(* IEC 61131-3 sources: daoli-st-library/DL_MathData (part 5) *)

(* ---- FC_DL_SaturateIncr.st ---- *)
(*==============================================================================
 * 组件名称 (Component)  : FC_DL_SaturateIncr
 * 所属子库 (Sublibrary) : DL_MathData ｜ 版本 (Version) : 1.0.0 ｜ 2026-11-23
 * 兼容性   (Platform)   : CODESYS 3.5+ / TwinCAT 3 / 汇川 InoProShop / 施耐德 Machine Expert
 *                         仅依赖 IEC 61131-3 算术运算符与 ABS，零厂商私有库
 * 功能描述 (Function)   : 带上下限的原地递增饱和（FC 形态）：把 VAR_IN_OUT 引脚 fX 原地
 *                         +1.0（步进常量 DL_SINC_STEP），结果超上限 fMax 则饱和到 fMax，
 *                         低于下限 fMin 则抬升到 fMin。用于配方号 / 档位 / 索引游标类
 *                         计数递增，替代任何不经限位的裸 `x := x + 1`。
 *                         **原地语义**：写回点唯一（段 5），返回 FALSE 的所有出口均不写 fX，
 *                         保证「失败不推进」。
 * 接口     (Interface)  : VAR_IN_OUT fX 被递增的量（本件原地更新）[工程单位]；
 *                         输入 fMin 下限、fMax 上限（有效域 fMin ≤ fMax）[工程单位]；
 *                         输出 fY 递增后值（镜像 fX）[工程单位]、bSaturated 本拍是否饱和、
 *                         eErrCode（E_DL_SaturateErr）；返回值 = 递增已生效标志。
 * 边界     (Boundary)   : ① fMin > fMax → 故障级 eBadLimit，fX 不写回（保持原值）。
 *                         ② 任一入参非有限 → 故障级 eNonFinite，fX 不写回。
 *                         ③ fX + 1 溢出为非有限 → 故障级 eNonFinite，fX 不写回（不饱和猜测）。
 *                         ④ 上限饱和与下限抬升为两个独立分支、两个独立码值（R190 归因唯一）。
 *                         ⑤ 容差 DL_SINC_EPS（1E-6）用于「恰好等于限值」的判定，禁浮点判等。
 *                         ⑥ 零全局耦合（无 GVL / VAR_EXTERNAL / 物理地址）。
 * 码表     (Codes)      : 本件不占用全局数字码位（R297 零码位范式）；出口为 BOOL + LREAL +
 *                         本文件内 enum E_DL_SaturateErr（全库唯一属主，与递减件共用同族枚举）。
 * 分工声明 (Scope)      : 递减同族件为 FC_DL_SaturateDecr（共用 E_DL_SaturateErr）；
 *                         整数类限位递增归 FC_DL_ClampDintChk 与 FC_DL_IndexClampEx。
 * 归属     (Ownership)  : E_DL_SaturateErr 归属本文件（全库唯一属主，R264）；
 *                         FC_DL_SaturateDecr 只引用不重声明。
 * 红线自检 (Redline)    : R1 ✓ 零 GVL ｜ R2 ✓ 零 %I/%Q ｜ R3 ✓ 纯 IEC ｜ R4 ✓ 非有限双判 +
 *                         上下限域闸 + 容差比较 ｜ R5 ✓ 逐行同行双语注释 ｜ R6 N/A（纯函数）
 *                         R7 N/A（无实例调用）
 * 修订历史 (Revision)   : 2026-11-23  v1.0.0  R78-B2 首版
 * 验收向量 (Acceptance) :
 *   A1 fX=4.0, fMin=0.0, fMax=10.0 → fX=5.0, fY=5.0, bSaturated=FALSE, eIncremented；
 *   A2 fX=10.0, fMin=0.0, fMax=10.0 → fX=10.0, bSaturated=TRUE, eSatHigh；
 *   A3 fX=9.5, fMin=0.0, fMax=10.0 → fX=10.0, bSaturated=TRUE, eSatHigh；
 *   A4 fX=-1.0, fMin=0.0, fMax=10.0 → fX=0.0, bSaturated=TRUE, eSatLow（抬升到下限）；
 *   A5 fX=5.0, fMin=10.0, fMax=0.0 → fX 保持 5.0, eBadLimit, 返回 FALSE。
 *============================================================================*)

(*-----------------------------------------------------------------------------
 * 枚举: E_DL_SaturateErr（递增 / 递减饱和出口码；信息级 = 0..9，故障级 = 10 起）
 *----------------------------------------------------------------------------*)
TYPE E_DL_SaturateErr :
(
    eIncremented := 0,   // 信息级：本拍在限内推进（递减件同样复用该成员）/ Info: advanced within limits
    eSatHigh     := 1,   // 信息级：上限饱和 / Info: saturated at the high limit
    eSatLow      := 2,   // 信息级：下限饱和（抬升到下限）/ Info: saturated at the low limit
    eBadLimit    := 10,  // 故障级：上下限倒置 / Fault: inverted limits
    eNonFinite   := 11   // 故障级：入参或结果非有限 / Fault: non-finite input or result
);
END_TYPE

FUNCTION FC_DL_SaturateIncr : BOOL
VAR_IN_OUT
    fX : LREAL;      // 被原地递增的量，成功时本件写回新值 [工程单位] / Value incremented in place, written back on success
END_VAR
VAR_INPUT
    fMin : LREAL;    // 下限 [工程单位] / Low limit in engineering unit
    fMax : LREAL;    // 上限，有效域 ≥ fMin [工程单位] / High limit in engineering unit, valid domain >= fMin
END_VAR
VAR_OUTPUT
    fY         : LREAL;             // 递增后值（镜像 fX）[工程单位] / Incremented value, mirror of fX
    bSaturated : BOOL;              // 本拍是否发生饱和 [-] / Saturation flag of this scan
    eErrCode   : E_DL_SaturateErr;  // 出口码 [-] / Outlet code
END_VAR
VAR
    _bBadX   : BOOL;   // fX 非有限标志 [-] / Non-finite flag of fX
    _bBadMin : BOOL;   // fMin 非有限标志 [-] / Non-finite flag of fMin
    _bBadMax : BOOL;   // fMax 非有限标志 [-] / Non-finite flag of fMax
    _fNext   : LREAL;  // 裸递增结果 = fX + 步进 [工程单位] / Raw incremented value before saturation
END_VAR
VAR CONSTANT
    DL_SINC_ZERO : LREAL := 0.0;     // 零基准 [-] / Zero base
    DL_SINC_ONE  : LREAL := 1.0;     // 递增步进常量 [-] / Increment step constant
    DL_SINC_EPS  : LREAL := 1.0E-6;  // 限值比较容差 [-] / Limit comparison tolerance
END_VAR

(* —— 段 0：出口预置安全侧 —— *)
FC_DL_SaturateIncr := FALSE;                         // 返回值预置未生效 / Return preset not applied
fY         := fX;                                    // 镜像出口取原值（失败不推进）/ Mirror keeps the original value on failure
bSaturated := FALSE;                                 // 饱和标志预清（单拍位统一预置）/ Single-shot flag preset
eErrCode   := E_DL_SaturateErr.eNonFinite;           // 预置最严码 / Preset strictest code

(* —— 段 1：入参非有限闸（R272 全量枚举 fX / fMin / fMax） —— *)
_bBadX   := (fX <> fX) OR ((fX - fX) <> DL_SINC_ZERO);                       // 被递增量非有限 / Value non-finite
_bBadMin := (fMin <> fMin) OR ((fMin - fMin) <> DL_SINC_ZERO);               // 下限非有限 / Low limit non-finite
_bBadMax := (fMax <> fMax) OR ((fMax - fMax) <> DL_SINC_ZERO);               // 上限非有限 / High limit non-finite
IF _bBadX OR _bBadMin OR _bBadMax THEN
    RETURN;                                          // 故障出口：fX 不写回 / Fault exit, fX not written
END_IF

(* —— 段 2：上下限域闸（倒置即组态缺陷，拒绝且不写回） —— *)
IF fMin > (fMax + DL_SINC_EPS) THEN
    eErrCode := E_DL_SaturateErr.eBadLimit;          // 故障级码 / Fault-level code
    RETURN;                                          // 返回 FALSE / Fault exit
END_IF

(* —— 段 3：裸递增与溢出复检 —— *)
_fNext := fX + DL_SINC_ONE;                          // 裸递增 / Raw increment
IF (_fNext <> _fNext) OR ((_fNext - _fNext) <> DL_SINC_ZERO) THEN
    eErrCode := E_DL_SaturateErr.eNonFinite;         // 故障级码：溢出为非有限 / Fault: overflow to non-finite
    RETURN;                                          // 返回 FALSE，fX 不写回 / Fault exit
END_IF

(* —— 段 4：上限饱和（独立分支 + 独立码值，R190） —— *)
IF _fNext > fMax THEN
    fY         := fMax;                              // 饱和到上限 / Saturate at the high limit
    fX         := fMax;                              // 原地写回（唯一写回点）/ Single write-back point
    bSaturated := TRUE;                              // 饱和标志 / Saturation flag
    eErrCode   := E_DL_SaturateErr.eSatHigh;         // 信息级：上限饱和 / Info: saturated high
    FC_DL_SaturateIncr := TRUE;                      // 递增已生效（饱和后值）/ Increment applied with saturation
    RETURN;
END_IF

(* —— 段 5：下限抬升（独立分支 + 独立码值，R190） —— *)
IF _fNext < fMin THEN
    fY         := fMin;                              // 抬升到下限 / Lift to the low limit
    fX         := fMin;                              // 原地写回（唯一写回点）/ Single write-back point
    bSaturated := TRUE;                              // 饱和标志 / Saturation flag
    eErrCode   := E_DL_SaturateErr.eSatLow;          // 信息级：下限饱和 / Info: saturated low
    FC_DL_SaturateIncr := TRUE;                      // 递增已生效（抬升后值）/ Increment applied with lift
    RETURN;
END_IF

(* —— 段 6：限内正常推进 —— *)
fY         := _fNext;                                // 正常推进结果 / Normal incremented value
fX         := _fNext;                                // 原地写回（唯一写回点）/ Single write-back point
bSaturated := FALSE;                                 // 未饱和 / Not saturated
eErrCode   := E_DL_SaturateErr.eIncremented;         // 信息级：限内推进 / Info: advanced within limits
FC_DL_SaturateIncr := TRUE;                          // 递增已生效 / Increment applied
END_FUNCTION

(* ---- FC_DL_SlewLimitLreal.st ---- *)
(*==============================================================================
 * 组件名称 (Component)  : FC_DL_SlewLimitLreal
 * 所属子库 (Sublibrary) : DL_MathData ｜ 版本 (Version) : 1.0.0 ｜ 2026-11-23
 * 兼容性   (Platform)   : CODESYS 3.5+ / TwinCAT 3 / 汇川 InoProShop / 施耐德 Machine Expert
 *                         仅依赖 IEC 61131-3 算术运算符、ABS 与标准转换函数，零厂商私有库
 * 功能描述 (Function)   : LREAL 精度斜率限幅（FC 形态）：与 FC_DL_RateLimitReal 同族，
 *                         但全链以 LREAL 计算，避免高精度位置 / 流量累加链在 REAL
 *                         单精度（约 7 位有效数字）上的步进量化误差。
 *                         **窄化出口**：fYReal 由 LREAL_TO_REAL 显式转换（R10），并在
 *                         超出 REAL 可表范围时饱和到 ±3.4028235E38 并置信息级
 *                         eNarrowClamp；窄化方向属于监护出口，饱和不放行是安全侧。
 *                         **契约声明**：fXPrev（VAR_IN_OUT）持有上一拍受限输出。
 * 接口     (Interface)  : 输入 fX 原始输入 [工程单位]、fRateMax 限幅速率 [单位/秒]、
 *                         fDt 采样周期 [s]；VAR_IN_OUT fXPrev 上一拍受限输出（本件写回，LREAL）；
 *                         输出 fY 限幅输出 [LREAL 工程单位]、fYReal 窄化出口 [REAL]、
 *                         eErrCode（E_DL_SlewLimitErr）；返回值 = 数值可信标志。
 * 边界     (Boundary)   : ① fRateMax ≤ 0 或 fDt ≤ 0 → 旁路，fY = fX（信息级 eBypass）。
 *                         ② 任一浮点入参非有限 → 故障级 eNonFinite，fY = 0 哨兵，返回 FALSE。
 *                         ③ 步进溢出为非有限 → 按旁路处理（信息级 eBypass）。
 *                         ④ 限幅后复检非有限 → 回退 fXPrev 并报故障。
 *                         ⑤ 窄化超 REAL 可表范围 → 饱和 + 信息级 eNarrowClamp（不改 LREAL 主出口）。
 *                         ⑥ 容差 DL_SLEW_EPS（1E-12，LREAL 口径；REAL 的 1E-6 在此过粗）。
 *                         ⑦ 零全局耦合（无 GVL / VAR_EXTERNAL / 物理地址）。
 * 码表     (Codes)      : 本件不占用全局数字码位（R297 零码位范式）；出口为 BOOL + LREAL +
 *                         本文件内 enum E_DL_SlewLimitErr（全库唯一属主）。
 * 分工声明 (Scope)      : REAL 精度同族件为 FC_DL_RateLimitReal；本件只做精度升级，
 *                         判据结构一致，便于同一工程内按量纲精度选型。
 * 归属     (Ownership)  : E_DL_SlewLimitErr 归属本文件（全库唯一属主，R264）。
 * 红线自检 (Redline)    : R1 ✓ 零 GVL ｜ R2 ✓ 零 %I/%Q ｜ R3 ✓ 纯 IEC ｜ R4 ✓ 非有限双判 +
 *                         容差比较 + 无除法 ｜ R5 ✓ 逐行同行双语注释 ｜ R6 N/A（纯函数）
 *                         R7 N/A（无实例调用） ｜ R10 ✓ LREAL_TO_REAL 显式窄化
 * 修订历史 (Revision)   : 2026-11-23  v1.0.0  R78-B2 首版
 * 验收向量 (Acceptance) :
 *   A1 fX=1.0, fPrev=0.0, fRateMax=0.1, fDt=1.0 → fY=0.1, fYReal=0.1, eLimited；
 *   A2 fX=1.0E-9, fPrev=0.0, fRateMax=1.0, fDt=1.0 → 增量在步进内 → fY=1.0E-9, eOk
 *      （REAL 精度件在同一向量上会因 1E-6 容差直通，本件用 1E-12 容差仍判直通但步进量可分辨）；
 *   A3 fX=5.0, fPrev=4.0, fRateMax=0.0, fDt=1.0 → 旁路 fY=5.0, eBypass, 返回 TRUE；
 *   A4 fX=NaN → fY=0.0, eNonFinite, 返回 FALSE；
 *   A5 fX=1.0E39（超 REAL 范围）, fPrev=0.0, fRateMax=1.0E40, fDt=1.0 → fY=1.0E39,
 *      fYReal=3.4028235E38（饱和）, eNarrowClamp。
 *============================================================================*)

(*-----------------------------------------------------------------------------
 * 枚举: E_DL_SlewLimitErr（LREAL 斜率限幅出口码；信息级 = 0..9，故障级 = 10 起）
 *----------------------------------------------------------------------------*)
TYPE E_DL_SlewLimitErr :
(
    eOk          := 0,   // 信息级：未超速，直通 / Info: within rate, pass-through
    eLimited     := 1,   // 信息级：本拍已按最大步进逼近 / Info: closed in by the max step this scan
    eBypass      := 2,   // 信息级：速率或周期越域，旁路输出原值 / Info: rate or period out of domain, bypassed
    ePrevRebuilt := 3,   // 信息级：fXPrev 未初始化或被污染，已重建 / Info: previous output rebuilt from fX
    eNarrowClamp := 4,   // 信息级：窄化出口超 REAL 可表范围，已饱和 / Info: narrowing saturated at REAL range
    eNonFinite   := 10   // 故障级：入参或结果非有限 / Fault: non-finite input or result
);
END_TYPE

FUNCTION FC_DL_SlewLimitLreal : BOOL
VAR_INPUT
    fX       : LREAL;   // 本拍原始输入 [工程单位，LREAL 精度] / Raw input this scan in engineering unit, LREAL precision
    fRateMax : LREAL;   // 允许最大变化速率，有效域 > 0 [单位/秒] / Max allowed rate, valid domain > 0 in unit per second
    fDt      : LREAL;   // 采样周期，有效域 > 0 [s] / Sampling period, valid domain > 0 in seconds
END_VAR
VAR_IN_OUT
    fXPrev : LREAL;     // 上一拍受限输出，本件写回新值 [工程单位] / Previous limited output, written back by this function
END_VAR
VAR_OUTPUT
    fY       : LREAL;              // 限幅输出（主出口，全精度）[工程单位] / Limited output, primary full-precision outlet
    fYReal   : REAL;               // 窄化出口（LREAL_TO_REAL 显式转换）[工程单位] / Narrowed outlet via explicit LREAL_TO_REAL
    eErrCode : E_DL_SlewLimitErr;   // 出口码 [-] / Outlet code
END_VAR
VAR
    _bBadX     : BOOL;    // fX 非有限标志 [-] / Non-finite flag of fX
    _bBadRate  : BOOL;    // fRateMax 非有限标志 [-] / Non-finite flag of fRateMax
    _bBadDt    : BOOL;    // fDt 非有限标志 [-] / Non-finite flag of fDt
    _bBadPrev  : BOOL;    // fXPrev 非有限标志 [-] / Non-finite flag of fXPrev
    _fMaxStep  : LREAL;   // 本拍允许最大步进 = fRateMax × fDt [工程单位] / Max step this scan
    _fDelta    : LREAL;   // 原始增量 = fX − fXPrev [工程单位] / Raw delta
    _fAbsDelta : LREAL;   // 增量绝对值 [工程单位] / Absolute delta
END_VAR
VAR CONSTANT
    DL_SLEW_ZERO  : LREAL := 0.0;              // 零基准与符号分界 [-] / Zero base and sign boundary
    DL_SLEW_EPS   : LREAL := 1.0E-12;          // LREAL 口径浮点同值判定容差 [-] / Float equality tolerance in LREAL terms
    DL_SLEW_RMAX  : LREAL := 3.4028235E38;     // REAL 正向可表上限（窄化饱和用） / Positive REAL maximum for narrowing saturation
    DL_SLEW_RNEG  : LREAL := -3.4028235E38;    // REAL 负向可表下限（窄化饱和用） / Negative REAL minimum for narrowing saturation
END_VAR

(* —— 段 0：出口预置安全侧 —— *)
FC_DL_SlewLimitLreal := FALSE;                       // 返回值预置不可信 / Return preset not trustworthy
fY      := DL_SLEW_ZERO;                             // LREAL 主出口哨兵 / Primary outlet sentinel
fYReal  := LREAL_TO_REAL(DL_SLEW_ZERO);              // 窄化出口哨兵（显式转换）/ Narrowed outlet sentinel via explicit conversion
eErrCode := E_DL_SlewLimitErr.eNonFinite;            // 预置最严码 / Preset strictest code

(* —— 段 1：入参非有限闸（R272 全量枚举 fX / fRateMax / fDt） —— *)
_bBadX    := (fX <> fX) OR ((fX - fX) <> DL_SLEW_ZERO);                          // fX 非有限 / fX non-finite
_bBadRate := (fRateMax <> fRateMax) OR ((fRateMax - fRateMax) <> DL_SLEW_ZERO);  // 速率非有限 / Rate non-finite
_bBadDt   := (fDt <> fDt) OR ((fDt - fDt) <> DL_SLEW_ZERO);                      // 周期非有限 / Period non-finite
IF _bBadX OR _bBadRate OR _bBadDt THEN
    RETURN;                                          // 故障出口：哨兵保持 / Fault exit, sentinels kept
END_IF

(* —— 段 2：上一拍输出有效性闸（未初始化或污染 → 以本拍输入重建） —— *)
_bBadPrev := (fXPrev <> fXPrev) OR ((fXPrev - fXPrev) <> DL_SLEW_ZERO);          // 前值非有限 / Previous value non-finite
IF _bBadPrev THEN
    fXPrev   := fX;                                  // 重建起点 / Rebuild the starting point
    eErrCode := E_DL_SlewLimitErr.ePrevRebuilt;      // 信息级：前值已重建 / Info: previous value rebuilt
END_IF

(* —— 段 3：速率 / 周期域闸（≤ 0 → 旁路，输出原 x） —— *)
IF (fRateMax <= DL_SLEW_ZERO) OR (fDt <= DL_SLEW_ZERO) THEN
    fY       := fX;                                  // 旁路输出原值 / Bypass keeps the raw input
    fXPrev   := fX;                                  // 前值同步 / Previous value follows
    eErrCode := E_DL_SlewLimitErr.eBypass;           // 信息级：旁路 / Info: bypassed
    fYReal   := LREAL_TO_REAL(fY);                   // 窄化出口同步（显式）/ Narrowed outlet follows
    FC_DL_SlewLimitLreal := TRUE;                    // 旁路输出可信 / Bypass output trustworthy
    RETURN;
END_IF

(* —— 段 4：本拍最大步进（乘后复检，溢出为旁路） —— *)
_fMaxStep := fRateMax * fDt;                         // 步进 = 速率 × 周期 / Step equals rate times period
IF (_fMaxStep <> _fMaxStep) OR ((_fMaxStep - _fMaxStep) <> DL_SLEW_ZERO) THEN
    fY       := fX;                                  // 步进不可表：放弃逼近 / Unrepresentable step: no approach
    fXPrev   := fX;                                  // 前值同步 / Previous value follows
    eErrCode := E_DL_SlewLimitErr.eBypass;           // 信息级：旁路 / Info: bypassed
    fYReal   := LREAL_TO_REAL(fY);                   // 窄化出口同步（显式）/ Narrowed outlet follows
    FC_DL_SlewLimitLreal := TRUE;                    // 原值可信 / Raw value trustworthy
    RETURN;
END_IF

(* —— 段 5：增量比较与逼近（上下行分列，R146） —— *)
_fDelta    := fX - fXPrev;                           // 原始增量 / Raw delta
_fAbsDelta := ABS(_fDelta);                          // 增量绝对值 / Absolute delta
IF _fAbsDelta <= (_fMaxStep + DL_SLEW_EPS) THEN
    fY       := fX;                                  // 未超速：直通 / Within rate: pass-through
    eErrCode := E_DL_SlewLimitErr.eOk;               // 信息级：正常 / Info: normal
ELSE
    IF _fDelta > DL_SLEW_ZERO THEN
        fY := fXPrev + _fMaxStep;                    // 上行逼近 / Approach upward
    ELSE
        fY := fXPrev - _fMaxStep;                    // 下行逼近 / Approach downward
    END_IF
    eErrCode := E_DL_SlewLimitErr.eLimited;          // 信息级：本拍受限 / Info: limited this scan
END_IF

(* —— 段 6：结果复检（非有限 → 回退前值并报故障） —— *)
IF (fY <> fY) OR ((fY - fY) <> DL_SLEW_ZERO) THEN
    fY       := fXPrev;                              // 回退上一有效值 / Fall back to the last valid value
    fYReal   := LREAL_TO_REAL(fY);                   // 窄化出口同步（显式）/ Narrowed outlet follows
    eErrCode := E_DL_SlewLimitErr.eNonFinite;        // 故障级码 / Fault-level code
    RETURN;                                          // 返回 FALSE / Fault exit
END_IF

(* —— 段 7：窄化出口（R10 显式转换 + 可表范围饱和 + 信息级声明） —— *)
IF fY > DL_SLEW_RMAX THEN
    fYReal := LREAL_TO_REAL(DL_SLEW_RMAX);           // 正向饱和 / Saturate positive
    eErrCode := E_DL_SlewLimitErr.eNarrowClamp;      // 信息级：窄化饱和 / Info: narrowing saturated
ELSIF fY < DL_SLEW_RNEG THEN
    fYReal := LREAL_TO_REAL(DL_SLEW_RNEG);           // 负向饱和 / Saturate negative
    eErrCode := E_DL_SlewLimitErr.eNarrowClamp;      // 信息级：窄化饱和 / Info: narrowing saturated
ELSE
    fYReal := LREAL_TO_REAL(fY);                     // 域内窄化（显式）/ In-range narrowing via explicit conversion
END_IF

fXPrev := fY;                                        // 前值写回（唯一写入点）/ Single write-back point
FC_DL_SlewLimitLreal := TRUE;                        // 输出可信 / Output trustworthy
END_FUNCTION

(* ---- FC_DL_SpeedUnitConvert.st ---- *)
// FC_DL_SpeedUnitConvert v1.0.0
// 开源溯源：brOscatLib / URL https://github.com/iec-oscat-mirror / 许可证 MIT / 借鉴 MS_TO_KMH 速度互转语义，clean-room 重写
(*
  道莅工业代码库 | DL_MathData | FC_DL_SpeedUnitConvert
  版本: 1.0.0 | 日期: 2026-11-23 | 轮次: R75
  功能: 速度单位双向互转 m/s ↔ km/h（eMode 选择方向），域闸防非有限与超量程
  邻件关系: 单位换算族 Temp/Press/Flow/Angle/Torque UnitConvert 的速度类补口；
            差异点：本件为线性比例换算（×3.6），温度族为仿射换算（含偏置），
            两者口径独立不共享码位（本件 16#0002_1901）
*)
TYPE E_DL_SpeedConvMode :
(
    eMsToKmh   := 0,   // m/s → km/h（乘 3.6）/ Meter per second to kilometer per hour
    eKmhToMs   := 1    // km/h → m/s（除以 3.6）/ Kilometer per hour to meter per second
);
END_TYPE

FUNCTION FC_DL_SpeedUnitConvert : REAL
VAR_INPUT
    fValue : REAL := 0.0;                        // 输入速度值 [m/s 或 km/h，随 eMode] / Input speed value
    eMode  : E_DL_SpeedConvMode := E_DL_SpeedConvMode.eMsToKmh;   // 换算方向选择 / Conversion direction selector
END_VAR
VAR_OUTPUT
    bValid   : BOOL;                             // 结果有效回执 [-] / Result validity receipt
    uErrorId : UDINT;                            // 事件码，0 = 无事件；16#0002_1901 = 输入非有限 / Event code
END_VAR
VAR CONSTANT
    DL_SPD_KMH_PER_MS : REAL := 3.6;             // 换算系数 1 m/s = 3.6 km/h [km/h per m/s] / Conversion factor
    DL_SPD_ABSMAX     : REAL := 1.0E12;          // 超量程闸（|v| 上限，防系数放大后溢出）[m/s|km/h] / Over-range gate
END_VAR

// —— 段 0：全路径缺省 —— //
bValid   := FALSE;                               // 有效回执预清 / Validity preset
uErrorId := 16#0000;                             // 事件码预清 / Event code preset
FC_DL_SpeedUnitConvert := 0.0;                   // 返回值缺省零 / Return default zero

// —— 段 1：非有限与超量程闸 —— //
IF (fValue <> fValue) OR (ABS(fValue) >= DL_SPD_ABSMAX) THEN   // NaN 自反 + 近 Inf 幅值闸 / NaN and magnitude gate
    uErrorId := 16#0002_1901;                    // 信息级：输入非有限或超量程（不置 bError） / Info level: invalid input
    RETURN;                                      // 返回零 / Return zero
END_IF

// —— 段 2：双向换算（CASE 全枚举 + ELSE 兜底） —— //
CASE eMode OF
E_DL_SpeedConvMode.eMsToKmh :                    // m/s → km/h / m/s to km/h
    FC_DL_SpeedUnitConvert := fValue * DL_SPD_KMH_PER_MS;    // ×3.6 / Multiply by 3.6
E_DL_SpeedConvMode.eKmhToMs :                    // km/h → m/s / km/h to m/s
    FC_DL_SpeedUnitConvert := fValue / DL_SPD_KMH_PER_MS;    // ÷3.6（常量非零，无除零风险）/ Divide by nonzero constant
ELSE                                             // 非法枚举兜底 / Illegal enum fallback
    uErrorId := 16#0002_1901;                    // 信息级：模式非法，返回零 / Info level: illegal mode
    RETURN;
END_CASE
bValid := TRUE;                                  // 有效回执 / Validity receipt
END_FUNCTION

(* ---- FC_DL_StatsMeanStdDev.st ---- *)
(*==============================================================================
 * 组件名称 (Component)  : FC_DL_StatsMeanStdDev
 * 所属子库 (Sublibrary) : DL_MathData
 * 当前版本 (Version)    : 1.0.0
 * 兼容性   (Platform)   : CODESYS 3.5+ / TwinCAT 3 / 汇川 InoProShop / 施耐德 Machine Expert
 *                         仅依赖 IEC 61131-3 标准数学（SQRT / ABS），零厂商私有库
 * 功能描述 (Function)   : 均值与标准差，采用 **Welford 单遍递推**（数值稳定、防溢出）：
 *                           k := k + 1
 *                           delta := x - mean
 *                           mean  := mean + delta / k
 *                           m2    := m2 + delta × (x - mean)
 *                         var := m2 / (k - 1)（样本方差，无偏），std := SQRT(var)。
 *                         相比「先求和再求平方和」的朴素两式算法，Welford 不会因
 *                         大均值配小方差发生灾难性抵消，也不要求预存全样本。
 *                         用途：称重一致性、加工尺寸波动、批次质量 SPC 判据输入。
 * 接口     (Interface)  : 输入 afSample 样本数组 [EU]、iCount 有效样本数 [个]（2..64）；
 *                         输出 fMean 均值 [EU]、fStdDev 样本标准差 [EU]、fVariance 样本方差 [EU^2]、
 *                         fSum 样本和 [EU]、bValid 结果可信标志、eErrCode（E_DL_StatsMsdErr）；
 *                         返回值 = bValid（TRUE = 三个统计量均可信）。
 * 边界     (Boundary)   : ① 属主边界：只算一阶/二阶统计量，不做离群剔除、不做分布检验。
 *                         ② 样本数域闸 2..64：<2 无样本方差定义（分母 k-1 = 0）→ 故障级 eBadCount，
 *                         **除零在结构上被排除**（先判点数后递推）。
 *                         ③ 非有限双判：全部参与计算的样本逐个枚举（i = 1..iCount），
 *                         任一非有限 → 故障级 eNonFinite（漏判单个样本会污染全部统计量）。
 *                         ④ 结果复检：mean / stddev / var 三者均做非有限复检；var 出现极小负值
 *                         （浮点舍入残差）→ 钳 0 并置信息级 eVarClamped，**不输出 NaN**。
 *                         ⑤ 零全局耦合（无 GVL / VAR_EXTERNAL / 物理地址）。
 * 分工声明 (Scope)      : 与 `FC_DL_StatsRmsCalc` 分工：RMS 含直流分量归那件、
 *                         均值+去均值标准差归本件；与 `FC_DL_StatsOutlierCount` 分工：
 *                         离群计数归那件（其内部自带 Welford，不跨件调用）。
 * 来源标签 (Source Tag) : 原创实现（无外部代码引入）
 * 码表     (Codes)      : 本件不占用全局数字码位；出口为 BOOL + 4×LREAL +
 *                         本文件内定义 enum E_DL_StatsMsdErr（全库唯一）。
 * 红线自检 (Redline)    : R1 ✓ 零 GVL/VAR_EXTERNAL ｜ R2 ✓ 零 %I/%Q/%M ｜ R3 ✓ 纯 IEC 61131-3
 *                         R4 ✓ 点数域闸（除零结构性排除）+ 全样本非有限双判 + 负方差钳位 ｜ R5 ✓ 声明逐行同行双语注释
 *                         R6 N/A（纯函数无状态机） ｜ R7 N/A（无实例调用）
 * 修订历史 (Revision)   : 2026-11-23  v1.0.0  R77 首版（批次 B3 · 序号 16）
 * 验收向量 (Acceptance) : ① afSample=[2,4,4,4,5,5,7,9], iCount=8 → fMean=5.0，
 *                         fVariance=32/7≈4.571428571，fStdDev≈2.138089935（容差 1E-6）；
 *                         ② afSample=[1,1,1], iCount=3 → fMean=1.0, fStdDev=0.0, eOk；
 *                         ③ iCount=1 → 返回 FALSE, eBadCount, fMean/fStdDev 哨兵 0；
 *                         ④ afSample[3]=NaN, iCount=8 → 返回 FALSE, eNonFinite；
 *                         ⑤ afSample=[10,10], iCount=2 → fMean=10.0, fVariance=0.0, fStdDev=0.0。
 *==============================================================================*)

(*-----------------------------------------------------------------------------
 * 枚举: E_DL_StatsMsdErr（均值/标准差统计错误码，归属 DL_MathData，与本件同文件，全库唯一属主）
 *----------------------------------------------------------------------------*)
TYPE E_DL_StatsMsdErr :
(
    eOk          := 0,   // 信息级：统计完成 / Info: statistics computed
    eVarClamped  := 1,   // 信息级：方差负残差已钳 0 / Info: negative variance residual clamped to zero
    eBadCount    := 2,   // 故障级：样本数越域 / Fault: sample count out of domain
    eNonFinite   := 3    // 故障级：样本含非有限值 / Fault: non-finite sample present
);
END_TYPE

FUNCTION FC_DL_StatsMeanStdDev : BOOL
VAR_INPUT
    afSample : ARRAY[1..64] OF LREAL;  // 样本数组 [EU] / Sample array
    iCount   : INT;                    // 有效样本数（2..64） [个] / Valid sample count, 2..64
END_VAR
VAR_OUTPUT
    fMean     : LREAL;  // 算术均值 [EU] / Arithmetic mean
    fStdDev   : LREAL;  // 样本标准差（分母 n-1） [EU] / Sample standard deviation
    fVariance : LREAL;  // 样本方差 [EU^2] / Sample variance
    fSum      : LREAL;  // 样本和（诊断用） [EU] / Sample sum for diagnostics
    bValid    : BOOL;   // 结果可信标志 [-] / Result trustworthy flag
    eErrCode  : E_DL_StatsMsdErr; // 错误码出口 [-] / Error code outlet
END_VAR
VAR
    _i       : INT;    // 样本遍历下标 [-] / Sample index
    _bNonFin : BOOL;   // 非有限标志 [-] / Non-finite flag
    _fMean   : LREAL;  // Welford 递推均值 [EU] / Recursive mean
    _fM2     : LREAL;  // Welford 二阶中心矩累加 [EU^2] / Second central moment accumulator
    _fDelta  : LREAL;  // 样本与当前均值之差 [EU] / Delta between sample and running mean
    _fSum    : LREAL;  // 样本和累加 [EU] / Sample sum accumulator
    _fVar    : LREAL;  // 方差（钳位前） [EU^2] / Variance before clamping
END_VAR
VAR CONSTANT
    DL_SMS_CNT_MIN : INT := 2;        // 样本数下限（n-1 必须 > 0） [个] / Count lower bound
    DL_SMS_CNT_MAX : INT := 64;       // 样本数上限（数组容量） [个] / Count upper bound
    DL_SMS_ZERO    : LREAL := 0.0;    // 零基准（含非有限判零） [-] / Zero base including non-finite probe
    DL_SMS_ONE     : LREAL := 1.0;    // 单位常数（Welford 分母 k-1 的基准） [-] / Unit constant
END_VAR

(* —— 段 0：出口预置安全值 —— *)
FC_DL_StatsMeanStdDev := FALSE;                    // 返回值预置无效 / Return preset invalid
fMean     := DL_SMS_ZERO;                          // 均值哨兵 / Mean sentinel
fStdDev   := DL_SMS_ZERO;                          // 标准差哨兵 / Standard deviation sentinel
fVariance := DL_SMS_ZERO;                          // 方差哨兵 / Variance sentinel
fSum      := DL_SMS_ZERO;                          // 样本和哨兵 / Sum sentinel
bValid    := FALSE;                                // 可信标志预置否 / Trust flag preset false
eErrCode  := E_DL_StatsMsdErr.eBadCount;           // 预置最严码 / Preset strictest code

(* —— 段 1：样本数域闸（先判点数，方差分母 n-1 的除零被结构性排除） —— *)
IF (iCount < DL_SMS_CNT_MIN) OR (iCount > DL_SMS_CNT_MAX) THEN
    RETURN;
END_IF

(* —— 段 2：非有限域闸（全部参与计算的样本逐项枚举） —— *)
_bNonFin := FALSE;
_i := 1;
WHILE _i <= iCount DO
    IF (afSample[_i] <> afSample[_i]) OR ((afSample[_i] - afSample[_i]) <> DL_SMS_ZERO) THEN
        _bNonFin := TRUE;                          // 样本非有限 / Sample non-finite
    END_IF
    _i := _i + 1;
END_WHILE
IF _bNonFin THEN
    eErrCode := E_DL_StatsMsdErr.eNonFinite;       // 故障级码 / Fault-level code
    RETURN;
END_IF

(* —— 段 3：Welford 单遍递推（数值稳定，防灾难性抵消与溢出） —— *)
_fMean := DL_SMS_ZERO;
_fM2   := DL_SMS_ZERO;
_fSum  := DL_SMS_ZERO;
_i     := 1;
WHILE _i <= iCount DO
    _fSum   := _fSum + afSample[_i];               // 样本和 / Sample sum
    _fDelta := afSample[_i] - _fMean;              // 与当前均值之差 / Delta from running mean
    _fMean  := _fMean + _fDelta / INT_TO_LREAL(_i);   // 均值更新（分母 i >= 1，无除零） / Mean update
    _fM2    := _fM2 + _fDelta * (afSample[_i] - _fMean);   // 二阶中心矩累加 / M2 accumulation
    _i := _i + 1;
END_WHILE

(* —— 段 4：方差与标准差（分母 n-1 已由段 1 保证 >= 1） —— *)
_fVar := _fM2 / INT_TO_LREAL(iCount - 1);          // 样本方差（无偏） / Unbiased sample variance
IF _fVar < DL_SMS_ZERO THEN
    _fVar    := DL_SMS_ZERO;                       // 浮点残差负值钳 0，绝不输出 NaN / Clamp residual negative
    eErrCode := E_DL_StatsMsdErr.eVarClamped;      // 信息级码 / Info code
ELSE
    eErrCode := E_DL_StatsMsdErr.eOk;              // 信息级成功 / Info success
END_IF
fStdDev := SQRT(_fVar);                            // 标准差（非负） / Standard deviation, non-negative

(* —— 段 5：结果复检（三个统计量逐一非有限复检） —— *)
IF (fStdDev <> fStdDev) OR (_fVar <> _fVar) OR (_fMean <> _fMean) THEN
    fMean     := DL_SMS_ZERO;                      // 复检异常全部回哨兵 / Recheck failed: all sentinels
    fStdDev   := DL_SMS_ZERO;
    fVariance := DL_SMS_ZERO;
    fSum      := DL_SMS_ZERO;
    eErrCode  := E_DL_StatsMsdErr.eNonFinite;      // 故障级码 / Fault-level code
    RETURN;
END_IF
IF (fStdDev < DL_SMS_ZERO) OR (_fVar < DL_SMS_ZERO) THEN
    fMean     := DL_SMS_ZERO;                      // 负统计量不可能，判内部不一致 / Negative statistics impossible
    fStdDev   := DL_SMS_ZERO;
    fVariance := DL_SMS_ZERO;
    fSum      := DL_SMS_ZERO;
    eErrCode  := E_DL_StatsMsdErr.eNonFinite;
    RETURN;
END_IF

(* —— 段 6：成功出口 —— *)
fMean     := _fMean;                               // 导出均值 / Export mean
fVariance := _fVar;                                // 导出方差 / Export variance
fSum      := _fSum;                                // 导出样本和 / Export sum
bValid    := TRUE;
FC_DL_StatsMeanStdDev := TRUE;                     // 统计可信 / Statistics trustworthy

END_FUNCTION

(* ---- FC_DL_StatsMinMaxWindow.st ---- *)
(*==============================================================================
 * 组件名称 (Component)  : FC_DL_StatsMinMaxWindow
 * 所属子库 (Sublibrary) : DL_MathData
 * 当前版本 (Version)    : 1.0.0
 * 兼容性   (Platform)   : CODESYS 3.5+ / TwinCAT 3 / 汇川 InoProShop / 施耐德 Machine Expert
 *                         仅依赖 IEC 61131-3 算术运算符，零厂商私有库
 * 功能描述 (Function)   : 窗口极值与发生时刻。在 afSample[1..iCount] 中找最小值与最大值，
 *                         并回传它们**首次出现**的位置下标与对应时刻（afStamp 为并行时刻表，
 *                         单位通常为相对秒 [s]）。并列时取**首次出现**（严格 < / > 比较），
 *                         行为确定可复现。
 *                         用途：压力峰值出现时刻、温度最低点定位、批次内极值-时刻归档、
 *                         配合趋势图做极值标注。
 * 接口     (Interface)  : 输入 afSample 样本数组 [EU]、afStamp 时刻表 [s]（与样本一一对应）、
 *                         iCount 有效样本数 [个]（1..64）；
 *                         输出 fMin 最小值 [EU]、fMax 最大值 [EU]、
 *                         iMinIndex / iMaxIndex 极值下标 [1..iCount]、
 *                         fMinStamp / fMaxStamp 极值时刻 [s]、
 *                         bValid 结果可信标志、eErrCode（E_DL_StatsMmErr）；
 *                         返回值 = bValid（TRUE = 六个出口量均可信）。
 * 边界     (Boundary)   : ① 属主边界：只取极值与时刻，不做滑动窗口跨周期保持（跨周期归 FB）、
 *                         不做极值个数统计。
 *                         ② 样本数域闸 1..64：1 点合法（min = max = 该点，下标 1）。
 *                         ③ 非有限双判：afSample 与 afStamp **两表**全部有效元素逐个枚举，
 *                         任一非有限 → 故障级 eNonFinite。只查样本表而漏查时刻表，
 *                         会让极值时刻静默变成 NaN 却被判「成功」。
 *                         ④ 全常量样本（min = max）合法：两下标同为首次出现位置。
 *                         ⑤ 时刻表不要求单调递增（允许环形缓冲乱序），本件不做序校验。
 *                         ⑥ 零全局耦合（无 GVL / VAR_EXTERNAL / 物理地址）。
 * 分工声明 (Scope)      : 与 `FC_DL_StatsMeanStdDev` 分工：一二阶矩归那件、极值归本件；
 *                         与 `FB_DL_PeakHoldFilter` 分工：跨周期峰值保持归那件、
 *                         单批窗口极值归本件。
 * 来源标签 (Source Tag) : 原创实现（无外部代码引入）
 * 码表     (Codes)      : 本件不占用全局数字码位；出口为 BOOL + 2×LREAL + 2×INT + 2×LREAL +
 *                         本文件内定义 enum E_DL_StatsMmErr（全库唯一）。
 * 红线自检 (Redline)    : R1 ✓ 零 GVL/VAR_EXTERNAL ｜ R2 ✓ 零 %I/%Q/%M ｜ R3 ✓ 纯 IEC 61131-3
 *                         R4 ✓ 点数域闸 + 双表全元素非有限双判 + 下标复检 ｜ R5 ✓ 声明逐行同行双语注释
 *                         R6 N/A（纯函数无状态机） ｜ R7 N/A（无实例调用）
 * 修订历史 (Revision)   : 2026-11-23  v1.0.0  R77 首版（批次 B3 · 序号 17）
 * 验收向量 (Acceptance) : ① afSample=[5,2,9,4], afStamp=[0,1,2,3], iCount=4 →
 *                         fMin=2.0（下标 2，时刻 1.0）, fMax=9.0（下标 3，时刻 2.0）, eOk；
 *                         ② afSample=[7,7,7], afStamp=[0,1,2], iCount=3 →
 *                         fMin=fMax=7.0，两下标均 1（首次出现）, 时刻均 0.0；
 *                         ③ iCount=0 → 返回 FALSE, eBadCount, 各出口哨兵 0；
 *                         ④ afStamp[2]=NaN, iCount=4 → 返回 FALSE, eNonFinite（漏查时刻表的反例）；
 *                         ⑤ iCount=1, afSample=[3.5], afStamp=[10.0] → fMin=fMax=3.5，时刻 10.0。
 *==============================================================================*)

(*-----------------------------------------------------------------------------
 * 枚举: E_DL_StatsMmErr（窗口极值统计错误码，归属 DL_MathData，与本件同文件，全库唯一属主）
 *----------------------------------------------------------------------------*)
TYPE E_DL_StatsMmErr :
(
    eOk        := 0,   // 信息级：统计完成 / Info: statistics computed
    eBadCount  := 1,   // 故障级：样本数越域 / Fault: sample count out of domain
    eNonFinite := 2,   // 故障级：样本或时刻含非有限值 / Fault: non-finite sample or stamp
    eInternal  := 9    // 故障级：极值下标越域（内部不一致） / Fault: extreme index out of domain
);
END_TYPE

FUNCTION FC_DL_StatsMinMaxWindow : BOOL
VAR_INPUT
    afSample : ARRAY[1..64] OF LREAL;  // 样本数组 [EU] / Sample array
    afStamp  : ARRAY[1..64] OF LREAL;  // 时刻表（与样本一一对应） [s] / Stamp table aligned with samples
    iCount   : INT;                    // 有效样本数（1..64） [个] / Valid sample count, 1..64
END_VAR
VAR_OUTPUT
    fMin      : LREAL;  // 最小值 [EU] / Minimum value
    fMax      : LREAL;  // 最大值 [EU] / Maximum value
    iMinIndex : INT;    // 最小值下标（首次出现） [1..iCount] / Minimum index, first occurrence
    iMaxIndex : INT;    // 最大值下标（首次出现） [1..iCount] / Maximum index, first occurrence
    fMinStamp : LREAL;  // 最小值发生时刻 [s] / Minimum stamp
    fMaxStamp : LREAL;  // 最大值发生时刻 [s] / Maximum stamp
    bValid    : BOOL;   // 结果可信标志 [-] / Result trustworthy flag
    eErrCode  : E_DL_StatsMmErr; // 错误码出口 [-] / Error code outlet
END_VAR
VAR
    _i         : INT;    // 样本遍历下标 [-] / Sample index
    _iMin      : INT;    // 最小值下标累计 [-] / Minimum index accumulator
    _iMax      : INT;    // 最大值下标累计 [-] / Maximum index accumulator
    _bNonFin   : BOOL;   // 非有限标志 [-] / Non-finite flag
    _fMin      : LREAL;  // 最小值累计 [EU] / Minimum accumulator
    _fMax      : LREAL;  // 最大值累计 [EU] / Maximum accumulator
END_VAR
VAR CONSTANT
    DL_SMM_CNT_MIN : INT := 1;        // 样本数下限 [个] / Count lower bound
    DL_SMM_CNT_MAX : INT := 64;       // 样本数上限（数组容量） [个] / Count upper bound
    DL_SMM_ZERO    : LREAL := 0.0;    // 零基准（含非有限判零） [-] / Zero base including non-finite probe
    DL_SMM_ONE     : INT := 1;        // 起始下标（IEC 1 基） [-] / Start index, IEC one-based
END_VAR

(* —— 段 0：出口预置安全值 —— *)
FC_DL_StatsMinMaxWindow := FALSE;                  // 返回值预置无效 / Return preset invalid
fMin      := DL_SMM_ZERO;                          // 最小值哨兵 / Minimum sentinel
fMax      := DL_SMM_ZERO;                          // 最大值哨兵 / Maximum sentinel
iMinIndex := 0;                                    // 最小值下标哨兵 / Minimum index sentinel
iMaxIndex := 0;                                    // 最大值下标哨兵 / Maximum index sentinel
fMinStamp := DL_SMM_ZERO;                          // 最小值时刻哨兵 / Minimum stamp sentinel
fMaxStamp := DL_SMM_ZERO;                          // 最大值时刻哨兵 / Maximum stamp sentinel
bValid    := FALSE;                                // 可信标志预置否 / Trust flag preset false
eErrCode  := E_DL_StatsMmErr.eBadCount;            // 预置最严码 / Preset strictest code

(* —— 段 1：样本数域闸 —— *)
IF (iCount < DL_SMM_CNT_MIN) OR (iCount > DL_SMM_CNT_MAX) THEN
    RETURN;
END_IF

(* —— 段 2：非有限域闸（样本表 + 时刻表双表逐项枚举） —— *)
_bNonFin := FALSE;
_i := 1;
WHILE _i <= iCount DO
    IF (afSample[_i] <> afSample[_i]) OR ((afSample[_i] - afSample[_i]) <> DL_SMM_ZERO) THEN
        _bNonFin := TRUE;                          // 样本非有限 / Sample non-finite
    END_IF
    IF (afStamp[_i] <> afStamp[_i]) OR ((afStamp[_i] - afStamp[_i]) <> DL_SMM_ZERO) THEN
        _bNonFin := TRUE;                          // 时刻非有限 / Stamp non-finite
    END_IF
    _i := _i + 1;
END_WHILE
IF _bNonFin THEN
    eErrCode := E_DL_StatsMmErr.eNonFinite;        // 故障级码 / Fault-level code
    RETURN;
END_IF

(* —— 段 3：极值扫描（严格比较 → 并列取首次出现） —— *)
_fMin  := afSample[DL_SMM_ONE];                    // 以首样本为初值 / Seed with first sample
_fMax  := afSample[DL_SMM_ONE];
_iMin  := DL_SMM_ONE;
_iMax  := DL_SMM_ONE;
_i     := 1;
WHILE _i <= iCount DO
    IF afSample[_i] < _fMin THEN
        _fMin := afSample[_i];                     // 更小值 / Smaller value
        _iMin := _i;
    END_IF
    IF afSample[_i] > _fMax THEN
        _fMax := afSample[_i];                     // 更大值 / Greater value
        _iMax := _i;
    END_IF
    _i := _i + 1;
END_WHILE

(* —— 段 4：下标复检（必须落在 1..iCount，否则判内部不一致） —— *)
IF (_iMin < DL_SMM_CNT_MIN) OR (_iMin > iCount) OR (_iMax < DL_SMM_CNT_MIN) OR (_iMax > iCount) THEN
    eErrCode := E_DL_StatsMmErr.eInternal;         // 故障级：下标越域 / Fault: index out of domain
    RETURN;
END_IF

(* —— 段 5：结果非有限复检（极值） —— *)
IF (_fMin <> _fMin) OR (_fMax <> _fMax) THEN
    eErrCode := E_DL_StatsMmErr.eNonFinite;
    RETURN;
END_IF

(* —— 段 6：成功出口（导出极值、下标与时刻） —— *)
fMin      := _fMin;
fMax      := _fMax;
iMinIndex := _iMin;
iMaxIndex := _iMax;
fMinStamp := afStamp[_iMin];                       // 极值时刻按下标回查 / Stamp looked up by index
fMaxStamp := afStamp[_iMax];
bValid    := TRUE;
eErrCode  := E_DL_StatsMmErr.eOk;                  // 信息级成功 / Info success
FC_DL_StatsMinMaxWindow := TRUE;                   // 统计可信 / Statistics trustworthy

END_FUNCTION

(* ---- FC_DL_StatsOutlierCount.st ---- *)
(*==============================================================================
 * 组件名称 (Component)  : FC_DL_StatsOutlierCount
 * 所属子库 (Sublibrary) : DL_MathData
 * 当前版本 (Version)    : 1.0.0
 * 兼容性   (Platform)   : CODESYS 3.5+ / TwinCAT 3 / 汇川 InoProShop / 施耐德 Machine Expert
 *                         仅依赖 IEC 61131-3 标准数学（ABS / SQRT），零厂商私有库
 * 功能描述 (Function)   : 离群点计数（3σ 判据）。步骤：
 *                         ① 用 Welford 单遍递推求均值与样本标准差（防溢出、防抵消）；
 *                         ② 逐点判 |x_i - mean| > fSigmaK × std，命中即计一个离群点；
 *                         ③ 回传离群个数、占比、判据阈值与两端样本值。
 *                         **样本不足保护**：样本数 < 8 时 σ 估计极不稳定（自由度过低），
 *                         本件不给出离群判定，回 iOutliers = 0、bValid = FALSE、
 *                         信息级码 eInsufficientSamples，让调用方明确知道「未判」而非「无离群」——
 *                         若静默返回 0，会被误当成「质量良好」。
 *                         **零离散保护**：std 近似 0（所有样本相同）时任何偏离都不可能存在，
 *                         回 0 并置信息级 eZeroSpread，避免 0 × k = 0 把全样本判成离群。
 * 接口     (Interface)  : 输入 afSample 样本数组 [EU]、iCount 有效样本数 [个]（2..64）、
 *                         fSigmaK 判据倍数（默认 3.0，必须 > 0） [倍]；
 *                         输出 iOutliers 离群点数 [个]、fOutlierRate 离群占比 [0..1]、
 *                         fMean 均值 [EU]、fStdDev 样本标准差 [EU]、fLimit 判定阈值带（k×σ） [EU]、
 *                         bValid 判定是否成立、eErrCode（E_DL_StatsOutErr）；
 *                         返回值 = bValid（**注意：样本不足时返回 FALSE**，与「无离群但判定成立」
 *                         严格区分——后者返回 TRUE 且 iOutliers = 0）。
 * 边界     (Boundary)   : ① 属主边界：只计数，不剔除、不替换离群点（剔除策略归调用方）。
 *                         ② 样本数域闸 2..64；< 8 判「样本不足」（信息级，返回 FALSE）。
 *                         ③ fSigmaK <= 0 → 故障级 eBadParam（0 倍会把全部样本判成离群）。
 *                         ④ 非有限双判：fSigmaK 与全部样本逐一枚举。
 *                         ⑤ 判据用严格大于（>），恰在边界上的点**不算**离群（保守口径，
 *                         避免阈值抖动导致计数跳变）。
 *                         ⑥ 零全局耦合（无 GVL / VAR_EXTERNAL / 物理地址）。
 * 分工声明 (Scope)      : 与 `FC_DL_StatsMeanStdDev` 分工：本件内部自带 Welford 以保持
 *                         单次调用语义（不跨件调用，避免多一次数组遍历与出口耦合）；
 *                         与 `FB_DL_HoldLastGoodFilter` 分工：坏值保持归那件。
 * 来源标签 (Source Tag) : 原创实现（无外部代码引入）
 * 码表     (Codes)      : 本件不占用全局数字码位；出口为 BOOL + INT + 5×LREAL +
 *                         本文件内定义 enum E_DL_StatsOutErr（全库唯一）。
 * 红线自检 (Redline)    : R1 ✓ 零 GVL/VAR_EXTERNAL ｜ R2 ✓ 零 %I/%Q/%M ｜ R3 ✓ 纯 IEC 61131-3
 *                         R4 ✓ 样本不足保护 + 零离散保护 + 倍数域闸 + 全样本非有限双判 ｜ R5 ✓ 声明逐行同行双语注释
 *                         R6 N/A（纯函数无状态机） ｜ R7 N/A（无实例调用）
 * 修订历史 (Revision)   : 2026-11-23  v1.0.0  R77 首版（批次 B3 · 序号 21）
 * 验收向量 (Acceptance) : ① afSample=[10,10,10,10,10,10,10,10,10,40], iCount=10, fSigmaK=3.0 →
 *                         mean=13.0, σ≈9.0（样本）；|40-13|=27 > 3×9.0≈27.0 边界 → 按严格 >
 *                         判定，27 与 27.0 相等时**不计**（保守）；取 fSigmaK=2.5 则计入 1 个；
 *                         ② afSample=[5,5,5,5,5,5,5,5], iCount=8, fSigmaK=3.0 →
 *                         std=0 → eZeroSpread，iOutliers=0，返回 TRUE；
 *                         ③ iCount=7 → 返回 FALSE, eInsufficientSamples（明确「未判」）；
 *                         ④ fSigmaK=0.0 → 返回 FALSE, eBadParam；
 *                         ⑤ iCount=0 → 返回 FALSE, eBadCount。
 *==============================================================================*)

(*-----------------------------------------------------------------------------
 * 枚举: E_DL_StatsOutErr（离群点统计错误码，归属 DL_MathData，与本件同文件，全库唯一属主）
 *----------------------------------------------------------------------------*)
TYPE E_DL_StatsOutErr :
(
    eOk                 := 0,   // 信息级：判定成立并完成计数 / Info: judgement valid and counted
    eZeroSpread         := 1,   // 信息级：零离散，无离群可能 / Info: zero spread, no outlier possible
    eInsufficientSamples:= 2,   // 信息级：样本不足 8 个，判定不成立 / Info: fewer than eight samples, judgement invalid
    eBadCount           := 3,   // 故障级：样本数越域 / Fault: sample count out of domain
    eNonFinite          := 4,   // 故障级：样本或倍数含非有限值 / Fault: non-finite sample or multiplier
    eBadParam           := 5    // 故障级：判据倍数非正 / Fault: non-positive sigma multiplier
);
END_TYPE

FUNCTION FC_DL_StatsOutlierCount : BOOL
VAR_INPUT
    afSample : ARRAY[1..64] OF LREAL;  // 样本数组 [EU] / Sample array
    iCount   : INT;                    // 有效样本数（2..64） [个] / Valid sample count, 2..64
    fSigmaK  : LREAL;                  // 判据倍数，必须 > 0，常取 3.0 [倍] / Sigma multiplier, must be positive
END_VAR
VAR_OUTPUT
    iOutliers    : INT;    // 离群点数 [个] / Outlier count
    fOutlierRate : LREAL;  // 离群占比 [0..1] / Outlier ratio
    fMean        : LREAL;  // 样本均值 [EU] / Sample mean
    fStdDev      : LREAL;  // 样本标准差 [EU] / Sample standard deviation
    fLimit       : LREAL;  // 判定阈值带 k×σ [EU] / Decision band width
    bValid       : BOOL;   // 判定是否成立 [-] / Whether the judgement is valid
    eErrCode     : E_DL_StatsOutErr; // 错误码出口 [-] / Error code outlet
END_VAR
VAR
    _i       : INT;    // 样本遍历下标 [-] / Sample index
    _iOut    : INT;    // 离群净额累加器（单点写入） [个] / Net outlier accumulator
    _bNonFin : BOOL;   // 非有限标志 [-] / Non-finite flag
    _fMean   : LREAL;  // Welford 递推均值 [EU] / Recursive mean
    _fM2     : LREAL;  // 二阶中心矩累加 [EU^2] / Second central moment accumulator
    _fDelta  : LREAL;  // 样本与均值之差 [EU] / Delta from running mean
    _fVar    : LREAL;  // 方差 [EU^2] / Variance
    _fStd    : LREAL;  // 标准差 [EU] / Standard deviation
    _fLimit  : LREAL;  // 判定带宽 k×σ [EU] / Decision band width
END_VAR
VAR CONSTANT
    DL_SOC_CNT_MIN  : INT := 2;        // 样本数下限 [个] / Count lower bound
    DL_SOC_CNT_MAX  : INT := 64;       // 样本数上限（数组容量） [个] / Count upper bound
    DL_SOC_CNT_STAT : INT := 8;        // 统计可信最小样本数 [个] / Minimum samples for a valid judgement
    DL_SOC_ZERO     : LREAL := 0.0;    // 零基准（含非有限判零） [-] / Zero base including non-finite probe
    DL_SOC_TINY     : LREAL := 1.0E-9; // 零离散判定阈值 [EU] / Zero-spread threshold
END_VAR

(* —— 段 0：出口预置安全值 —— *)
FC_DL_StatsOutlierCount := FALSE;                  // 返回值预置无效（判定未成立） / Return preset invalid
iOutliers    := 0;                                 // 离群计数哨兵 / Outlier count sentinel
fOutlierRate := DL_SOC_ZERO;                       // 离群占比哨兵 / Outlier ratio sentinel
fMean        := DL_SOC_ZERO;                       // 均值哨兵 / Mean sentinel
fStdDev      := DL_SOC_ZERO;                       // 标准差哨兵 / Standard deviation sentinel
fLimit       := DL_SOC_ZERO;                       // 判定带哨兵 / Decision band sentinel
bValid       := FALSE;                             // 判定成立标志预置否 / Judgement valid preset false
eErrCode     := E_DL_StatsOutErr.eBadCount;        // 预置最严码 / Preset strictest code

(* —— 段 1：样本数域闸 —— *)
IF (iCount < DL_SOC_CNT_MIN) OR (iCount > DL_SOC_CNT_MAX) THEN
    RETURN;
END_IF

(* —— 段 2：非有限域闸（倍数 + 全部样本逐项枚举） —— *)
_bNonFin := (fSigmaK <> fSigmaK) OR ((fSigmaK - fSigmaK) <> DL_SOC_ZERO);
_i := 1;
WHILE _i <= iCount DO
    IF (afSample[_i] <> afSample[_i]) OR ((afSample[_i] - afSample[_i]) <> DL_SOC_ZERO) THEN
        _bNonFin := TRUE;
    END_IF
    _i := _i + 1;
END_WHILE
IF _bNonFin THEN
    eErrCode := E_DL_StatsOutErr.eNonFinite;       // 故障级码 / Fault-level code
    RETURN;
END_IF

(* —— 段 3：判据倍数域闸（必须严格为正，否则全部样本都会被判离群） —— *)
IF fSigmaK <= DL_SOC_ZERO THEN
    eErrCode := E_DL_StatsOutErr.eBadParam;        // 故障级：倍数非正 / Fault: non-positive multiplier
    RETURN;
END_IF

(* —— 段 4：Welford 单遍求均值与标准差（样本不足时也先算出来供诊断） —— *)
_fMean := DL_SOC_ZERO;
_fM2   := DL_SOC_ZERO;
_i     := 1;
WHILE _i <= iCount DO
    _fDelta := afSample[_i] - _fMean;
    _fMean  := _fMean + _fDelta / INT_TO_LREAL(_i);            // 分母 i >= 1，无除零 / Denominator at least one
    _fM2    := _fM2 + _fDelta * (afSample[_i] - _fMean);
    _i := _i + 1;
END_WHILE
_fVar := _fM2 / INT_TO_LREAL(iCount - 1);          // 样本方差（n-1 已由段 1 保证 >= 1） / Unbiased variance
IF _fVar < DL_SOC_ZERO THEN
    _fVar := DL_SOC_ZERO;                          // 浮点残差负值钳 0 / Clamp residual negative
END_IF
_fStd := SQRT(_fVar);                              // 标准差 / Standard deviation
fMean   := _fMean;                                 // 导出均值（诊断量，任何分支都可信） / Export mean
fStdDev := _fStd;                                  // 导出标准差 / Export standard deviation

(* —— 段 5：样本不足保护（< 8 个不判，明确回「未判」而非「无离群」） —— *)
IF iCount < DL_SOC_CNT_STAT THEN
    iOutliers    := 0;
    fOutlierRate := DL_SOC_ZERO;
    fLimit       := DL_SOC_ZERO;
    bValid       := FALSE;                         // 判定不成立 / Judgement invalid
    eErrCode     := E_DL_StatsOutErr.eInsufficientSamples;   // 信息级：样本不足 / Info: insufficient samples
    FC_DL_StatsOutlierCount := FALSE;              // 返回 FALSE 与「成立且 0 离群」严格区分 / Distinguish from valid zero
    RETURN;
END_IF

(* —— 段 6：零离散保护（所有样本相同，无离群可能） —— *)
IF _fStd < DL_SOC_TINY THEN
    iOutliers    := 0;
    fOutlierRate := DL_SOC_ZERO;
    fLimit       := DL_SOC_ZERO;
    bValid       := TRUE;                          // 判定成立：确实无离群 / Judgement valid: truly no outlier
    eErrCode     := E_DL_StatsOutErr.eZeroSpread;  // 信息级：零离散 / Info: zero spread
    FC_DL_StatsOutlierCount := TRUE;
    RETURN;
END_IF

(* —— 段 7：离群计数（严格大于判据带，恰在边界不计） —— *)
_fLimit := fSigmaK * _fStd;                        // 判定带宽 k×σ / Decision band width
fLimit  := _fLimit;
_iOut   := 0;
_i      := 1;
WHILE _i <= iCount DO
    IF ABS(afSample[_i] - _fMean) > _fLimit THEN
        _iOut := _iOut + 1;                        // 命中离群（单点累加） / Count one outlier
    END_IF
    _i := _i + 1;
END_WHILE
iOutliers    := _iOut;                             // 导出离群数 / Export outlier count
fOutlierRate := INT_TO_LREAL(_iOut) / INT_TO_LREAL(iCount);   // 占比（分母 n >= 8，无除零） / Ratio

(* —— 段 8：结果复检（非有限 + 计数域） —— *)
IF (fLimit <> fLimit) OR (fMean <> fMean) OR (fStdDev <> fStdDev) THEN
    iOutliers    := 0;
    fOutlierRate := DL_SOC_ZERO;
    fLimit       := DL_SOC_ZERO;
    bValid       := FALSE;
    eErrCode     := E_DL_StatsOutErr.eNonFinite;
    RETURN;
END_IF
IF (_iOut < 0) OR (_iOut > iCount) THEN
    iOutliers    := 0;
    fOutlierRate := DL_SOC_ZERO;
    bValid       := FALSE;
    eErrCode     := E_DL_StatsOutErr.eBadCount;
    RETURN;
END_IF

(* —— 段 9：成功出口 —— *)
bValid   := TRUE;
eErrCode := E_DL_StatsOutErr.eOk;                  // 信息级成功 / Info success
FC_DL_StatsOutlierCount := TRUE;                   // 判定成立且计数可信 / Judgement valid and count trustworthy

END_FUNCTION

(* ---- FC_DL_StatsPercentile.st ---- *)
(*==============================================================================
 * 组件名称 (Component)  : FC_DL_StatsPercentile
 * 所属子库 (Sublibrary) : DL_MathData
 * 当前版本 (Version)    : 1.0.0
 * 兼容性   (Platform)   : CODESYS 3.5+ / TwinCAT 3 / 汇川 InoProShop / 施耐德 Machine Expert
 *                         仅依赖 IEC 61131-3 标准数学（TRUNC / MIN / MAX），零厂商私有库
 * 功能描述 (Function)   : 分位数计算（P50 / P90 / P95 等），排序法 + 线性插值。
 *                         ① 把有效样本复制到内部缓冲（**不改写调用方数组**）；
 *                         ② 冒泡排序升序（N <= 64，最坏 64×63/2 = 2016 次比较，单拍可接受）；
 *                         ③ 位置 pos := (p/100) × (n - 1)（0 基）；
 *                            lo := TRUNC(pos)，frac := pos - lo；
 *                            结果 := buf[lo] × (1 - frac) + buf[lo+1] × frac。
 *                         取整一律用 TRUNC 后按余量插值，**不使用 TRUNC(x)+1 这类手工进位**
 *                         （R 加固清单要求：向上取整禁止 TRUNC+1，须先 TRUNC 再按余量进位）。
 * 接口     (Interface)  : 输入 afSample 样本数组 [EU]、iCount 有效样本数 [个]（1..64）、
 *                         fPercent 百分位 [%]（0..100，0 = 最小，100 = 最大）；
 *                         输出 fResult 分位数值 [EU]、fPos 位置（0 基，诊断用）[-]、
 *                         bInterpolated 是否发生两点插值、bValid 结果可信、
 *                         eErrCode（E_DL_StatsPctErr）；
 *                         返回值 = bValid。
 * 边界     (Boundary)   : ① 属主边界：只算单个分位点；P50/P90/P95 由调用方三次调用
 *                         （避免本件内部固定三个出口，保持通用）。
 *                         ② 样本数域闸 1..64；越域 → 故障级 eBadCount。n=1 时 pos 恒 0，结果即唯一值。
 *                         ③ 百分位域闸 0..100；越域 → 故障级 eBadPercent（不做静默钳位，
 *                         避免把「配置写错 950」当成 95 用）。
 *                         ④ 非有限双判：全部有效样本逐项枚举。
 *                         ⑤ 插值上界保护：lo 若达到 n-1（pos 恰为最大值）则退化为单点取值，
 *                         不读 buf[lo+1]（**杜绝数组越界**）。
 *                         ⑥ 零全局耦合（无 GVL / VAR_EXTERNAL / 物理地址）。
 * 分工声明 (Scope)      : 与 `FC_DL_StatsMeanStdDev` 分工：矩统计归那件、序统计归本件；
 *                         与 `FC_DL_StatsOutlierCount` 分工：离群计数归那件。
 * 来源标签 (Source Tag) : 原创实现（无外部代码引入）
 * 码表     (Codes)      : 本件不占用全局数字码位；出口为 BOOL + 2×LREAL + BOOL +
 *                         本文件内定义 enum E_DL_StatsPctErr（全库唯一）。
 * 红线自检 (Redline)    : R1 ✓ 零 GVL/VAR_EXTERNAL ｜ R2 ✓ 零 %I/%Q/%M ｜ R3 ✓ 纯 IEC 61131-3
 *                         R4 ✓ 点数/百分位双域闸 + 全样本非有限双判 + 插值下标越界保护 ｜ R5 ✓ 声明逐行同行双语注释
 *                         R6 N/A（纯函数无状态机） ｜ R7 N/A（无实例调用）
 * 修订历史 (Revision)   : 2026-11-23  v1.0.0  R77 首版（批次 B3 · 序号 18）
 * 验收向量 (Acceptance) : ① afSample=[1,2,3,4,5], iCount=5, fPercent=50 → pos=0.5×4=2.0,
 *                         lo=2, frac=0 → fResult=3.0（一点起算：buf[3]=3.0）, bInterpolated=FALSE；
 *                         ② 同上, fPercent=90 → pos=0.9×4=3.6, lo=3, frac=0.6 →
 *                         fResult=4×0.4+5×0.6=4.6（容差 1E-9）, bInterpolated=TRUE；
 *                         ③ 同上, fPercent=100 → pos=4 → 退化单点 → fResult=5.0（不越界）；
 *                         ④ fPercent=101 → 返回 FALSE, eBadPercent；
 *                         ⑤ iCount=0 → 返回 FALSE, eBadCount。
 *==============================================================================*)

(*-----------------------------------------------------------------------------
 * 枚举: E_DL_StatsPctErr（分位数统计错误码，归属 DL_MathData，与本件同文件，全库唯一属主）
 *----------------------------------------------------------------------------*)
TYPE E_DL_StatsPctErr :
(
    eOk          := 0,   // 信息级：分位数计算完成 / Info: percentile computed
    eBadCount    := 1,   // 故障级：样本数越域 / Fault: sample count out of domain
    eBadPercent  := 2,   // 故障级：百分位越域（0..100） / Fault: percentile out of range
    eNonFinite   := 3,   // 故障级：样本含非有限值 / Fault: non-finite sample present
    eInternal    := 9    // 故障级：插值下标越界（内部不一致） / Fault: interpolation index out of range
);
END_TYPE

FUNCTION FC_DL_StatsPercentile : BOOL
VAR_INPUT
    afSample : ARRAY[1..64] OF LREAL;  // 样本数组（只读） [EU] / Sample array, read-only
    iCount   : INT;                    // 有效样本数（1..64） [个] / Valid sample count, 1..64
    fPercent : LREAL;                  // 百分位 [%]（0..100） / Percentile in percent
END_VAR
VAR_OUTPUT
    fResult       : LREAL;  // 分位数值 [EU] / Percentile value
    fPos          : LREAL;  // 插值位置（0 基，诊断用） [-] / Interpolation position, zero-based
    bInterpolated : BOOL;   // 是否发生两点插值 [-] / Whether two-point interpolation occurred
    bValid        : BOOL;   // 结果可信标志 [-] / Result trustworthy flag
    eErrCode      : E_DL_StatsPctErr; // 错误码出口 [-] / Error code outlet
END_VAR
VAR
    _afBuf     : ARRAY[1..64] OF LREAL;  // 内部排序缓冲（不改写调用方数组） [EU] / Internal sort buffer
    _i         : INT;    // 外层遍历下标 [-] / Outer index
    _j         : INT;    // 内层遍历下标 [-] / Inner index
    _iLo       : INT;    // 位置下整（0 基） [-] / Floor index, zero-based
    _diLo      : DINT;   // 下整中间量（LREAL→DINT，再收窄到 INT） [-] / Floor intermediate, LREAL to DINT then INT
    _bNonFin   : BOOL;   // 非有限标志 [-] / Non-finite flag
    _bSwapped  : BOOL;   // 冒泡交换标志 [-] / Bubble swap flag
    _fTmp      : LREAL;  // 交换临时量 [EU] / Swap temporary
    _fPosR     : LREAL;  // 位置（0 基） [-] / Position, zero-based
    _fFrac     : LREAL;  // 位置小数部分（余量） [-] / Fractional remainder
END_VAR
VAR CONSTANT
    DL_SPC_CNT_MIN : INT := 1;        // 样本数下限 [个] / Count lower bound
    DL_SPC_CNT_MAX : INT := 64;       // 样本数上限（数组容量） [个] / Count upper bound
    DL_SPC_PCT_MIN : LREAL := 0.0;    // 百分位下限 [%] / Percentile lower bound
    DL_SPC_PCT_MAX : LREAL := 100.0;  // 百分位上限 [%] / Percentile upper bound
    DL_SPC_ZERO    : LREAL := 0.0;    // 零基准（含非有限判零） [-] / Zero base including non-finite probe
    DL_SPC_ONE     : LREAL := 1.0;    // 单位常数 [-] / Unit constant
    DL_SPC_HUND    : LREAL := 100.0;  // 百分数换算因子 [-] / Percent scaling factor
    DL_SPC_ONE_I   : INT := 1;        // 下标单位（IEC 1 基） [-] / Index unit, IEC one-based
END_VAR

(* —— 段 0：出口预置安全值 —— *)
FC_DL_StatsPercentile := FALSE;                    // 返回值预置无效 / Return preset invalid
fResult       := DL_SPC_ZERO;                      // 结果哨兵 / Result sentinel
fPos          := DL_SPC_ZERO;                      // 位置哨兵 / Position sentinel
bInterpolated := FALSE;                            // 插值标志预置否 / Interpolation preset false
bValid        := FALSE;                            // 可信标志预置否 / Trust flag preset false
eErrCode      := E_DL_StatsPctErr.eBadCount;       // 预置最严码 / Preset strictest code

(* —— 段 1：样本数域闸 —— *)
IF (iCount < DL_SPC_CNT_MIN) OR (iCount > DL_SPC_CNT_MAX) THEN
    RETURN;
END_IF

(* —— 段 2：百分位域闸（越域不做静默钳位，避免配置错误被掩盖） —— *)
IF (fPercent <> fPercent) OR (fPercent < DL_SPC_PCT_MIN) OR (fPercent > DL_SPC_PCT_MAX) THEN
    eErrCode := E_DL_StatsPctErr.eBadPercent;      // 故障级：百分位越域 / Fault: percentile out of range
    RETURN;
END_IF

(* —— 段 3：非有限域闸（全部有效样本逐项枚举） —— *)
_bNonFin := FALSE;
_i := 1;
WHILE _i <= iCount DO
    IF (afSample[_i] <> afSample[_i]) OR ((afSample[_i] - afSample[_i]) <> DL_SPC_ZERO) THEN
        _bNonFin := TRUE;
    END_IF
    _i := _i + 1;
END_WHILE
IF _bNonFin THEN
    eErrCode := E_DL_StatsPctErr.eNonFinite;       // 故障级码 / Fault-level code
    RETURN;
END_IF

(* —— 段 4：复制到内部缓冲（不改写调用方数组，R 纪律） —— *)
FOR _i := DL_SPC_ONE_I TO iCount DO
    _afBuf[_i] := afSample[_i];
END_FOR;

(* —— 段 5：冒泡排序升序（N <= 64，比较次数有界） —— *)
FOR _i := 1 TO (iCount - 1) DO
    _bSwapped := FALSE;
    FOR _j := 1 TO (iCount - _i) DO
        IF _afBuf[_j] > _afBuf[_j + DL_SPC_ONE_I] THEN
            _fTmp                := _afBuf[_j];
            _afBuf[_j]           := _afBuf[_j + DL_SPC_ONE_I];
            _afBuf[_j + 1]       := _fTmp;
            _bSwapped            := TRUE;          // 本趟发生交换 / Swap happened in this pass
        END_IF
    END_FOR;
    IF NOT _bSwapped THEN
        _i := iCount;                              // 已有序：提前收敛（仍受 FOR 上界约束） / Early convergence
    END_IF
END_FOR;

(* —— 段 6：位置计算（0 基，先 TRUNC 再按余量插值，禁 TRUNC+1 手工进位） —— *)
_fPosR := (fPercent / DL_SPC_HUND) * INT_TO_LREAL(iCount - 1);   // pos = (p/100)*(n-1)
fPos   := _fPosR;
_diLo  := LREAL_TO_DINT(TRUNC(_fPosR));            // 先 TRUNC 再转整（禁 TRUNC+1 手工进位） / Truncate then convert
_iLo   := DINT_TO_INT(_diLo);                      // 收窄到 INT（0..63，越界由下两段钳位） / Narrow to INT
IF _iLo < 0 THEN
    _iLo := 0;                                     // 下标下限保护 / Lower index guard
END_IF
IF _iLo > (iCount - 1) THEN
    _iLo := iCount - 1;                            // 下标上限保护 / Upper index guard
END_IF
_fFrac := _fPosR - INT_TO_LREAL(_iLo);             // 余量（0..1） / Remainder
IF _fFrac < DL_SPC_ZERO THEN
    _fFrac := DL_SPC_ZERO;
END_IF
IF _fFrac > DL_SPC_ONE THEN
    _fFrac := DL_SPC_ONE;
END_IF

(* —— 段 7：取值（插值上界保护：lo 达末位时退化为单点，杜绝越界） —— *)
IF _iLo >= (iCount - 1) THEN
    fResult       := _afBuf[iCount];               // 末位单点取值 / Single-point value at the tail
    bInterpolated := FALSE;
ELSE
    fResult := _afBuf[_iLo + DL_SPC_ONE_I] * (DL_SPC_ONE - _fFrac)
             + _afBuf[_iLo + 1 + DL_SPC_ONE_I] * _fFrac;   // 两点线性插值 / Two-point linear interpolation
    bInterpolated := TRUE;
END_IF

(* —— 段 8：结果复检（非有限 + 落在 [min, max] 闭包内） —— *)
IF (fResult <> fResult) OR ((fResult - fResult) <> DL_SPC_ZERO) THEN
    fResult       := DL_SPC_ZERO;
    bInterpolated := FALSE;
    eErrCode      := E_DL_StatsPctErr.eNonFinite;
    RETURN;
END_IF
IF (fResult < _afBuf[DL_SPC_ONE_I]) OR (fResult > _afBuf[iCount]) THEN
    fResult       := DL_SPC_ZERO;                  // 越出样本闭包：内部不一致 / Outside sample envelope
    bInterpolated := FALSE;
    eErrCode      := E_DL_StatsPctErr.eInternal;
    RETURN;
END_IF

(* —— 段 9：成功出口 —— *)
bValid   := TRUE;
eErrCode := E_DL_StatsPctErr.eOk;                  // 信息级成功 / Info success
FC_DL_StatsPercentile := TRUE;                     // 分位数可信 / Percentile trustworthy

END_FUNCTION

(* ---- FC_DL_StatsZeroCrossRate.st ---- *)
(*==============================================================================
 * 组件名称 (Component)  : FC_DL_StatsZeroCrossRate
 * 所属子库 (Sublibrary) : DL_MathData
 * 当前版本 (Version)    : 1.0.0
 * 兼容性   (Platform)   : CODESYS 3.5+ / TwinCAT 3 / 汇川 InoProShop / 施耐德 Machine Expert
 *                         仅依赖 IEC 61131-3 算术运算符，零厂商私有库
 * 功能描述 (Function)   : 过零率统计（振动 / 流量脉动的频域粗特征）。
 *                         以 fThreshold（通常为 0，也可取样本均值作「过均值率」）为基准，
 *                         逐点比较相对阈值的位置（+1 = 高于阈值，-1 = 低于阈值，0 = 恰等于），
 *                         统计**位置符号发生翻转**的次数（双向翻转合并为单一净额计数）。
 *                         恰等于阈值的样本**不改变当前符号**（跳过而非计为新符号），
 *                         避免直流偏置或量化平台把翻转数虚增。
 *                         过零率 = 翻转数 / (n - 1)，即相邻样本对的翻转比例 [0..1]；
 *                         频率近似 ≈ 过零率 × 采样率 / 2（本件不回传频率，仅回传比例，
 *                         时基由调用方掌握）。
 * 接口     (Interface)  : 输入 afSample 样本数组 [EU]、iCount 有效样本数 [个]（2..64）、
 *                         fThreshold 判定阈值 [EU]（通常 0）；
 *                         输出 iCrossings 翻转次数 [次]、fRate 翻转比例 [0..1]、
 *                         fRatePercent 翻转百分比 [%]、bValid 结果可信、
 *                         eErrCode（E_DL_StatsZcrErr）；
 *                         返回值 = bValid。
 * 边界     (Boundary)   : ① 属主边界：只统计翻转比例，不换算 Hz（缺时基）、不做频谱分析。
 *                         ② 样本数域闸 2..64：n=1 时「相邻对」不存在，翻转率无定义 → 故障级 eBadCount
 *                         （除零防护：分母 n-1 必须 >= 1）。
 *                         ③ 非有限双判：**fThreshold 与全部样本逐一枚举**（漏判阈值会让
 *                         整个符号判定静默退化）。
 *                         ④ 全样本恰等于阈值（符号始终未定）→ 翻转数 0、比例 0.0、
 *                         置信息级 eNoSignDefined（不是故障：数据确实无方向信息）。
 *                         ⑤ 双向翻转合并为单一累加器 iCrossings（不分别计数后相加，
 *                         避免两处写入不一致）。
 *                         ⑥ 零全局耦合（无 GVL / VAR_EXTERNAL / 物理地址）。
 * 分工声明 (Scope)      : 与 `FC_DL_StatsRmsCalc` 分工：幅值特征归那件、翻转特征归本件；
 *                         与 `FB_DL_StatsZeroCrossRate`（若后续入库的跨周期件）分工：
 *                         本件为单批窗口统计，无跨周期状态。
 * 来源标签 (Source Tag) : 原创实现（无外部代码引入）
 * 码表     (Codes)      : 本件不占用全局数字码位；出口为 BOOL + INT + 2×LREAL +
 *                         本文件内定义 enum E_DL_StatsZcrErr（全库唯一）。
 * 红线自检 (Redline)    : R1 ✓ 零 GVL/VAR_EXTERNAL ｜ R2 ✓ 零 %I/%Q/%M ｜ R3 ✓ 纯 IEC 61131-3
 *                         R4 ✓ 点数域闸（分母 n-1 除零排除）+ 阈值与样本非有限双判 + 单点写入 ｜ R5 ✓ 声明逐行同行双语注释
 *                         R6 N/A（纯函数无状态机） ｜ R7 N/A（无实例调用）
 * 修订历史 (Revision)   : 2026-11-23  v1.0.0  R77 首版（批次 B3 · 序号 20）
 * 验收向量 (Acceptance) : ① afSample=[1,-1,1,-1], iCount=4, fThreshold=0 → 翻转 3 次,
 *                         fRate=3/3=1.0, fRatePercent=100.0, eOk, TRUE；
 *                         ② afSample=[1,2,3,4], iCount=4, fThreshold=0 → 翻转 0 次, fRate=0.0；
 *                         ③ afSample=[1,0,-1], iCount=3, fThreshold=0 → 符号 +1 → 跳过 → -1，
 *                         翻转 1 次（零值未计新符号）, fRate=0.5；
 *                         ④ afSample=[0,0,0], fThreshold=0 → 翻转 0 次, eNoSignDefined（信息级）；
 *                         ⑤ iCount=1 → 返回 FALSE, eBadCount（分母 n-1 会为 0）。
 *==============================================================================*)

(*-----------------------------------------------------------------------------
 * 枚举: E_DL_StatsZcrErr（过零率统计错误码，归属 DL_MathData，与本件同文件，全库唯一属主）
 *----------------------------------------------------------------------------*)
TYPE E_DL_StatsZcrErr :
(
    eOk            := 0,   // 信息级：统计完成 / Info: computed
    eNoSignDefined := 1,   // 信息级：样本全部等于阈值，无符号信息 / Info: all samples equal threshold
    eBadCount      := 2,   // 故障级：样本数越域（n-1 会为 0） / Fault: sample count out of domain
    eNonFinite     := 3    // 故障级：阈值或样本含非有限值 / Fault: non-finite threshold or sample
);
END_TYPE

FUNCTION FC_DL_StatsZeroCrossRate : BOOL
VAR_INPUT
    afSample   : ARRAY[1..64] OF LREAL;  // 样本数组 [EU] / Sample array
    iCount     : INT;                    // 有效样本数（2..64） [个] / Valid sample count, 2..64
    fThreshold : LREAL;                  // 判定阈值（通常 0） [EU] / Decision threshold, usually zero
END_VAR
VAR_OUTPUT
    iCrossings  : INT;    // 符号翻转次数 [次] / Number of sign flips
    fRate       : LREAL;  // 翻转比例（翻转数 / (n-1)） [0..1] / Flip ratio
    fRatePercent: LREAL;  // 翻转百分比 [%] / Flip percentage
    bValid      : BOOL;   // 结果可信标志 [-] / Result trustworthy flag
    eErrCode    : E_DL_StatsZcrErr; // 错误码出口 [-] / Error code outlet
END_VAR
VAR
    _i        : INT;    // 样本遍历下标 [-] / Sample index
    _iPrev    : INT;    // 上一有效符号（+1 / -1 / 0 = 未定） [-] / Previous sign, zero means undetermined
    _iCur     : INT;    // 当前符号 [-] / Current sign
    _iCross   : INT;    // 翻转净额累加器（单点写入） [次] / Net flip accumulator, single point
    _bNonFin  : BOOL;   // 非有限标志 [-] / Non-finite flag
    _fRate    : LREAL;  // 比例（钳位前） [-] / Ratio before clamping
END_VAR
VAR CONSTANT
    DL_SZC_CNT_MIN : INT := 2;        // 样本数下限（相邻对至少一对） [个] / Count lower bound
    DL_SZC_CNT_MAX : INT := 64;       // 样本数上限（数组容量） [个] / Count upper bound
    DL_SZC_HUND    : LREAL := 100.0;  // 百分数换算因子 [-] / Percent scaling factor
    DL_SZC_ZERO    : LREAL := 0.0;    // 零基准（含非有限判零） [-] / Zero base including non-finite probe
    DL_SZC_ONE     : LREAL := 1.0;    // 比例上限 [-] / Ratio upper bound
    DL_SZC_SIGN_P  : INT := 1;        // 符号：高于阈值 / Sign above threshold
    DL_SZC_SIGN_N  : INT := -1;       // 符号：低于阈值 / Sign below threshold
    DL_SZC_SIGN_0  : INT := 0;        // 符号：未定（恰等于阈值） / Sign undetermined
END_VAR

(* —— 段 0：出口预置安全值 —— *)
FC_DL_StatsZeroCrossRate := FALSE;                 // 返回值预置无效 / Return preset invalid
iCrossings   := 0;                                 // 翻转计数哨兵 / Flip count sentinel
fRate        := DL_SZC_ZERO;                       // 比例哨兵 / Ratio sentinel
fRatePercent := DL_SZC_ZERO;                       // 百分比哨兵 / Percentage sentinel
bValid       := FALSE;                             // 可信标志预置否 / Trust flag preset false
eErrCode     := E_DL_StatsZcrErr.eBadCount;        // 预置最严码 / Preset strictest code

(* —— 段 1：样本数域闸（分母 n-1 必须 >= 1，除零结构性排除） —— *)
IF (iCount < DL_SZC_CNT_MIN) OR (iCount > DL_SZC_CNT_MAX) THEN
    RETURN;
END_IF

(* —— 段 2：非有限域闸（阈值 + 全部样本逐项枚举） —— *)
_bNonFin := (fThreshold <> fThreshold) OR ((fThreshold - fThreshold) <> DL_SZC_ZERO);
_i := 1;
WHILE _i <= iCount DO
    IF (afSample[_i] <> afSample[_i]) OR ((afSample[_i] - afSample[_i]) <> DL_SZC_ZERO) THEN
        _bNonFin := TRUE;                          // 样本非有限 / Sample non-finite
    END_IF
    _i := _i + 1;
END_WHILE
IF _bNonFin THEN
    eErrCode := E_DL_StatsZcrErr.eNonFinite;       // 故障级码 / Fault-level code
    RETURN;
END_IF

(* —— 段 3：符号翻转扫描（恰等于阈值不改符号；双向翻转合并为单一累加器） —— *)
_iPrev  := DL_SZC_SIGN_0;                          // 符号未定 / Sign undetermined
_iCross := 0;
_i      := 1;
WHILE _i <= iCount DO
    IF afSample[_i] > fThreshold THEN
        _iCur := DL_SZC_SIGN_P;                    // 高于阈值 / Above threshold
    ELSIF afSample[_i] < fThreshold THEN
        _iCur := DL_SZC_SIGN_N;                    // 低于阈值 / Below threshold
    ELSE
        _iCur := DL_SZC_SIGN_0;                    // 恰等于阈值：本点不定义符号 / Undetermined at threshold
    END_IF

    IF _iCur <> DL_SZC_SIGN_0 THEN
        IF (_iPrev <> DL_SZC_SIGN_0) AND (_iCur <> _iPrev) THEN
            _iCross := _iCross + 1;                // 符号翻转一次（单点写入） / One flip
        END_IF
        _iPrev := _iCur;                           // 更新有效符号 / Update effective sign
    END_IF
    _i := _i + 1;
END_WHILE

(* —— 段 4：翻转比例（分母 n-1 >= 1，已由段 1 保证） —— *)
_fRate := INT_TO_LREAL(_iCross) / INT_TO_LREAL(iCount - 1);   // 翻转比例 / Flip ratio
_fRate := MIN(MAX(_fRate, DL_SZC_ZERO), DL_SZC_ONE);         // 显式约束 0..1 / Constrain 0..1
fRate        := _fRate;
fRatePercent := _fRate * DL_SZC_HUND;              // 百分比 / Percentage
iCrossings   := _iCross;

(* —— 段 5：无符号信息判定（全样本等于阈值） —— *)
IF _iPrev = DL_SZC_SIGN_0 THEN
    eErrCode := E_DL_StatsZcrErr.eNoSignDefined;   // 信息级：无方向信息 / Info: no directional information
ELSE
    eErrCode := E_DL_StatsZcrErr.eOk;              // 信息级成功 / Info success
END_IF

(* —— 段 6：结果复检（非有限 + 计数非负 + 不超相邻对数） —— *)
IF (fRate <> fRate) OR (fRatePercent <> fRatePercent) THEN
    iCrossings   := 0;
    fRate        := DL_SZC_ZERO;
    fRatePercent := DL_SZC_ZERO;
    eErrCode     := E_DL_StatsZcrErr.eNonFinite;
    RETURN;
END_IF
IF (iCrossings < 0) OR (iCrossings > (iCount - 1)) THEN
    iCrossings   := 0;                             // 计数越界：内部不一致 / Count out of range
    fRate        := DL_SZC_ZERO;
    fRatePercent := DL_SZC_ZERO;
    eErrCode     := E_DL_StatsZcrErr.eBadCount;
    RETURN;
END_IF

(* —— 段 7：成功出口 —— *)
bValid := TRUE;
FC_DL_StatsZeroCrossRate := TRUE;                  // 统计可信 / Statistics trustworthy

END_FUNCTION

(* ---- FC_DL_StdDevOnline.st ---- *)
(*==============================================================================
 * 组件名称 (Component)  : FC_DL_StdDevOnline
 * 所属子库 (Sublibrary) : DL_MathData
 * 当前版本 (Version)    : 1.0.0
 * 兼容性   (Platform)   : CODESYS 3.5+ / TwinCAT 3 / 汇川 InoProShop / 施耐德 Machine Expert
 *                         仅依赖 Standard.library（SQRT），零厂商私有库
 * 功能描述 (Function)   : Welford 单遍在线标准差（数值稳定型，免"先求和再减均方"的灾难性抵消）。
 *                         每次调用吞入一个样本，就地更新调用方持有的累加器 ST_DL_WelfordAcc：
 *                           nCount ← nCount + 1
 *                           fDelta  ← x − fMean
 *                           fMean   ← fMean + fDelta / nCount
 *                           fDelta2 ← x − fMean（注意用的是**更新后**的均值）
 *                           fM2     ← fM2 + fDelta × fDelta2
 *                         样本标准差 s = SQRT(fM2 / (nCount − 1))，返回 LREAL。
 * 无状态边界 (Stateless): **本 FC 自身零内部状态**（IEC 61131-3 的 FC 不得持有静态变量，本件遵守）。
 *                         全部跨拍状态由调用方通过 VAR_IN_OUT 累加器 stAcc 持有——这意味着：
 *                         ① 一个累加器实例 = 一路数据流，多路统计必须各用各的累加器（严禁共用）；
 *                         ② 调用方可在任意时刻把 stAcc 清零来重开统计窗（本件不提供隐式清零）；
 *                         ③ 本 FC 可重入、可并发、可放在任何 POU 内调用，结果只取决于入参与 stAcc。
 *                         若调用方希望"封装成自持状态的块"，请在外层包一层 FB 持有该累加器，
 *                         而不要把状态藏进本 FC（那会破坏无状态契约）。
 * 接口     (Interface)  : 入 fSample 新样本、stAcc 累加器（VAR_IN_OUT，读改写）；出 bValid 有效
 *                         （nCount >= 2 且样本有限）、fMean 当前均值、fM2 平方和、fStdDev 返回。
 * 边界     (Boundary)   : ① nCount < 2 → 标准差无定义，返回 0.0 且 bValid=FALSE（**不作 0 语义**
 *                         ——调用方必须查 bValid 才可用该值）；② 非有限样本（NaN/Inf，用 x<>x 自反
 *                         判 NaN、（x−x）<>(x−x) 判 Inf）→ 不入累加器、返回上次可用值域外的 0.0、
 *                         bValid=FALSE、bNonFin=TRUE——污染源绝不进状态，否则均值被永久毒化；
 *                         ③ fM2 累加可能因浮点误差出极小负值 → 开方前钳到 0（防 SQRT 负参得 NaN）；
 *                         ④ nCount 达上限 DL_WELFORD_MAX_N（16#00FF_FFFF）后不再自增，bSaturated=TRUE，
 *                         返回当前标准差（防 UDINT 回绕把 nCount 归零导致除零）。
 * 依赖     (Depends)    : 无 DL_ 内部依赖（仅本文件内的 ST_DL_WelfordAcc）；标准库仅 SQRT
 * 来源标签 (Source Tag) : T2-1 ◐（公开经典算法 Welford 1962 单遍方差；ST 重写 + 防御包装，零代码行复制）
 * 码表     (Codes)      : 本件不占用任何全局数字码位。异常出口为 BOOL（bValid / bNonFin /
 *                         bSaturated）；数字码位待主控收口阶段统一派号。
 * 红线自检 (Redline)    : R1 ✓ 零 GVL/VAR_EXTERNAL ｜ R2 ✓ 零 %I/%Q/%M ｜ R3 ✓ 纯 IEC 61131-3
 *                         R4 ✓ n<2 防除零 + 非有限闸 + 负方差钳位 ｜ R5 ✓ 声明逐行同行双语注释
 *                         R6 N/A（无状态机） ｜ R7 N/A（无实例调用）
 * 修订历史 (Revision)   : 2026-11-19  v1.0.0  R46 首版（批次 1 · 序号 5）
 *==============================================================================*)

TYPE ST_DL_WelfordAcc :
STRUCT
    nCount : UDINT := 0;    // 已吞入样本数（调用方所有，须初值 0） [个] / Samples consumed, caller-owned, init 0
    fMean  : LREAL := 0.0;  // 当前均值 μ [工程单位] / Running mean [engineering unit]
    fM2    : LREAL := 0.0;  // 均值偏差平方和 Σ(x−μ)² [工程单位²] / Sum of squared deviations [unit squared]
END_STRUCT
END_TYPE

FUNCTION FC_DL_StdDevOnline : LREAL
VAR_INPUT
    fSample : LREAL := 0.0;    // 本拍新样本（非有限样本被拒收） [工程单位] / New sample this scan, non-finite samples rejected
END_VAR
VAR_IN_OUT
    stAcc : ST_DL_WelfordAcc;  // 累加器（调用方持有，本 FC 零内部状态） [混合] / Accumulator owned by caller, this FC holds no state
END_VAR
VAR_OUTPUT
    bValid     : BOOL;         // 标准差有效（nCount >= 2 且本拍样本被接收或历史可用） [-] / StdDev valid
    bNonFin    : BOOL;         // 本拍样本非有限，已被拒收（未污染累加器） [-] / Sample non-finite and rejected
    bSaturated : BOOL;         // 样本数已达上限，停止自增（防 UDINT 回绕） [-] / Sample count capped
    fMean      : LREAL;        // 当前均值（出口镜像，便于 HMI 直读） [工程单位] / Mean mirror for HMI
    fM2        : LREAL;        // 当前平方和（出口镜像） [工程单位²] / M2 mirror
END_VAR
VAR
    fDelta  : LREAL;           // x − 旧均值 [工程单位] / Sample minus old mean
    fDelta2 : LREAL;           // x − 新均值 [工程单位] / Sample minus new mean
    fVar    : LREAL;           // 样本方差（分母 n−1） [工程单位²] / Sample variance with n-1 denominator
END_VAR
VAR CONSTANT
    DL_WELFORD_MAX_N : UDINT := 16#00FF_FFFF;   // 样本数上限，留足余量防回绕 [个] / Sample cap with wrap margin
    DL_WELFORD_ZERO  : LREAL := 0.0;            // 零基准（负方差钳位用） [无量纲] / Zero baseline for variance clamping
END_VAR

(* —— 段 1：出口初始化（任何路径下返回值确定） —— *)
FC_DL_StdDevOnline := 0.0;      // 缺省返回 0.0，须配 bValid 才可用 / Default 0.0, meaningful only with bValid
bValid     := FALSE;            // 先假定无效 / Assume invalid
bNonFin    := FALSE;            // 非有限标志清零 / Non-finite flag cleared
bSaturated := FALSE;            // 饱和标志清零 / Saturation flag cleared

(* —— 段 2：非有限闸（污染源不入状态，否则均值被永久毒化） —— *)
bNonFin := (fSample <> fSample)                             // NaN 自反判（判等禁令唯一例外） / NaN self-reflexive test
        OR ((fSample - fSample) <> (fSample - fSample));    // Inf 判：Inf−Inf 得 NaN，NaN≠NaN 为真 / Inf test via Inf minus Inf
IF bNonFin THEN
    fMean := stAcc.fMean;           // 回放当前均值，不改状态 / Replay mean without touching state
    fM2   := stAcc.fM2;             // 回放当前平方和 / Replay M2
    bValid := stAcc.nCount >= 2;    // 历史可用的前提下仍报有效（本拍未参与） / Still valid from history, sample excluded
    IF bValid THEN
        IF stAcc.nCount >= 2 THEN
            fVar := stAcc.fM2 / UDINT_TO_LREAL(stAcc.nCount - 1);    // 分母 n−1，n>=2 已闸 / n-1 denominator, guarded by n>=2
            IF fVar < DL_WELFORD_ZERO THEN
                fVar := DL_WELFORD_ZERO;                             // 负方差钳位（浮点误差） / Clamp negative variance
            END_IF
            FC_DL_StdDevOnline := SQRT(fVar);                        // 返回历史标准差 / Return historical StdDev
        END_IF
    END_IF
    RETURN;                         // 提前返回，累加器未被触碰 / Early return, accumulator untouched
END_IF

(* —— 段 3：样本数上限闸（防 UDINT 回绕把 nCount 归零） —— *)
IF stAcc.nCount >= DL_WELFORD_MAX_N THEN
    bSaturated := TRUE;                     // 达上限 / Cap reached
    fMean := stAcc.fMean;                   // 回放 / Replay
    fM2   := stAcc.fM2;                     // 回放 / Replay
    fVar  := stAcc.fM2 / UDINT_TO_LREAL(stAcc.nCount - 1);   // 上限远大于 2，分母安全 / Cap far above 2, denominator safe
    IF fVar < DL_WELFORD_ZERO THEN
        fVar := DL_WELFORD_ZERO;            // 负方差钳位 / Clamp
    END_IF
    FC_DL_StdDevOnline := SQRT(fVar);       // 返回当前标准差（不再更新） / Return current StdDev, no further update
    bValid := TRUE;                         // 历史统计仍有效 / Historical statistics still valid
    RETURN;
END_IF

(* —— 段 4：Welford 单遍更新（就地写回调用方累加器） —— *)
stAcc.nCount := stAcc.nCount + 1;                                   // 计数自增（已过上限闸） / Increment count, cap already gated
fDelta       := fSample - stAcc.fMean;                              // x − 旧均值 / Sample minus old mean
stAcc.fMean  := stAcc.fMean + (fDelta / UDINT_TO_LREAL(stAcc.nCount));   // 均值增量更新，分母 >= 1 恒安全 / Mean update, denominator >= 1
fDelta2      := fSample - stAcc.fMean;                              // x − 新均值 / Sample minus updated mean
stAcc.fM2    := stAcc.fM2 + (fDelta * fDelta2);                     // M2 累加（Welford 核心式） / M2 accumulation

(* —— 段 5：出口映射（n<2 无定义，返回 0 且 bValid=FALSE） —— *)
fMean := stAcc.fMean;               // 均值出口 / Mean outlet
fM2   := stAcc.fM2;                 // 平方和出口 / M2 outlet
IF stAcc.nCount >= 2 THEN
    fVar := stAcc.fM2 / UDINT_TO_LREAL(stAcc.nCount - 1);   // 样本方差（分母 n−1） / Sample variance
    IF fVar < DL_WELFORD_ZERO THEN
        fVar := DL_WELFORD_ZERO;                            // 负方差钳位（浮点误差不可开方） / Clamp negative variance
    END_IF
    FC_DL_StdDevOnline := SQRT(fVar);                       // 标准差 / Standard deviation
    bValid := TRUE;                                         // 有效 / Valid
ELSE
    FC_DL_StdDevOnline := 0.0;                              // 单样本无离散度，返回 0 但标无效 / Single sample: 0 but invalid
    bValid := FALSE;
END_IF

END_FUNCTION

(* ---- FC_DL_StringToDint.st ---- *)
(*
    组件名称 : FC_DL_StringToDint
    所属子库 : DL_MathData
    当前版本 : 1.0.2
    兼 容 性 : CODESYS V3.5+ / TwinCAT 3 / 汇川 InoProShop；仅依赖 Standard.library
    功能描述 : 整数字符串严格解析，补 FC_DL_StringToLReal 的整数族缺口（配方号 / 站号 / 批次号）。
              取舍 ①：不委托任何平台串转数值内建 —— 三家平台对非法字符、前导空格、符号重复的处理各不相同，
              有的返回 0、有的抛异常、有的静默截断，且都不告诉调用方错在第几位；现场最贵的不是「失败」，
              而是「成功但值不对」。本件逐字符推进，判断口径完全一致，并给出首个非法字符位置。
              取舍 ②：升位到 LINT 累加，每步先判界再落账 —— DINT 域中间量在 214748364 × 10 + 9 处已越界，
              直接在 DINT 里累加必然回绕；LINT 域足够宽，判界判的是 LINT 与 DINT 上下界的比较，安全。
              取舍 ③：负域上界取 2147483648 而非 2147483647 —— DINT_MIN 的绝对值比 DINT_MAX 大 1，
              用同一个上界会把 "-2147483648" 误判溢出（有符号整数边界必须双侧分开写，禁单侧 ABS 判据）。
              取舍 ④：溢出后返回「夹到边界」的值并置 bValid = FALSE —— 夹域值便于现场看出「方向对了但超了」，
              比返回 0 更容易定位问题；同时绝不把夹域值当有效值输出。
    开源溯源 : 原创实现（T0-5/T0-6 变体线）。字符判定与位置报错口径与库内 FC_DL_StringToLReal 同源，；本件为 IEC 61131-3 标准语义的道莅防御性实现（原创实现，零外部源码复制）。
              但字符集、累加类型、溢出判据全部按整数域重写。无外部源码参考，码位与分级 100% 自有。
    本文件内含 : FUNCTION FC_DL_StringToDint（单 POU）
                 同文件 TYPE E_DL_StrToDintState（归属本子库，全库唯一）
    依 赖 : 无 DL_ 内部依赖；Standard.library: LEN / MID / FIND
    红线自检 : R1 ✓ 零全局变量与外部变量 ｜ R2 ✓ 零物理 IO 地址
              R3 ✓ 纯 IEC 61131-3 ｜ R4 ✓ 空串闸 + 非法字符定位 + 双侧溢出判界 + WHILE 守卫计数器
              R5 ✓ 全变量中英双语同行注释 ｜ R6 ✓ ENUM + CASE + ELSE 兜底（非法状态落 038C）
              R7 N/A 无定时器、无沿检测实例 ｜ R8 ✓ 上下界、长度上限、守卫上限全常量化
    错误码   : 16#0001_0448 [信息级] 前后空格已忽略，解析正常，bValid = TRUE
               16#0001_0449 [信息级] 预留禁用（不得挪用）
               16#0001_038A [故障级] 空串或仅符号，nErrPos = 长度 + 1，返回 0，bValid = FALSE
               16#0001_038B [故障级] 数值溢出，返回夹到边界的值，bValid = FALSE，bError = TRUE（R41 P0-3 配对补齐）
               16#0001_038C [故障级] 非法字符（含 CASE 落 ELSE 的非法状态兜底，不新占码位），返回 0，bValid = FALSE
    码位总账 : 16#0001_0448 用 / 16#0001_0449 预留 ｜ 16#0001_038A 用 / 16#0001_038B 用 / 16#0001_038C 用
    遗留假设 : ① MID 参数序按 IEC 标准为 MID(串, 长度, 位置)，库内既有件同序；若某平台改为 MID(串, 位置, 长度)，
              本件会取到错字符 —— 属已知平台差异，须在编译门槛里核对（现有库内 9 处用法同序，风险已收敛）。
              ② FIND 返回 1 基位置、未命中返回 0，为 Standard.library 口径推导，未逐平台实测。
              ③ 字符串比较只用 = 与 <>，不用 < / >（部分平台未实现 STRING 排序比较），故数字字符判定走 FIND 表查。
    修订历史 :
        2026-11-16  v1.0.0  首版，R21 批次 3 入库
        2026-11-16  v1.0.1  R21 终审修复（轻微）：溢出分支原先只置 bOverflow / bAbort，未写 nErrPos，
                            导致 eErr = 038B（故障级）与 nErrPos = 0（「无错」哨兵）并存，现场按位置
                            指向排错时会得到「有故障但无位置」的矛盾诊断。现溢出位与非法字符位同口径
                            写入 nErrPos。对外引脚契约、返回值夹域策略、码位均不变。
        2026-11-19  v1.0.2  R41 P0-3 返修（R40 发现）：段 4 溢出出口 eErr := 16#0001_038B 原未
                            配对 bError := TRUE（R101 配对缺失），故障级码静默。现赋值行 3 行内
                            显式补配对置位，码表同步登记。VERSION/MANUAL 同步升级。
*)

(*-----------------------------------------------------------------------------
 * 枚举: E_DL_StrToDintState（归属本函数，与其同文件发布，全库唯一）
 * 含义: 逐字符解析的四态推进，成员值写死便于工程持久化
 *----------------------------------------------------------------------------*)
TYPE E_DL_StrToDintState :
(
    eLeadSpace := 0,    // 前导空格态：跳空格，遇非空格转符号态 / leading blank state, moves to the sign state on any other character
    eSign      := 10,   // 符号态：取前导正负号或直接进数字态 / sign state, consumes the leading sign or falls through to the digits
    eDigits    := 20,   // 数字态：逐位累加，遇尾随空格转结束态 / digits state, accumulates and moves to done on a trailing blank
    eDone      := 30    // 结束态：只允许尾随空格，别的字符一律非法 / done state, only trailing blanks are accepted
);
END_TYPE

FUNCTION FC_DL_StringToDint : DINT
VAR_INPUT
    sIn             : STRING;          // 待解析文本，最长 255 字符，允许前后空格 [字符] / input text, up to 255 characters, blanks allowed on both ends [char]
    bAllowSign      : BOOL := TRUE;    // 是否允许前导 +/− 号 / whether a leading sign is allowed
END_VAR
VAR_OUTPUT
    eErr            : UDINT;           // 错误码，0=正常；16#0001_04XX 信息级 / 16#0001_03XX 故障级 / error id, 0=ok
    bError          : BOOL;            // 故障级标志，eErr 落 16#0001_03XX 时为 TRUE / fault flag, TRUE on fault-level eErr
    bValid          : BOOL;            // 返回值是否可用 / result usable flag
    nErrPos         : INT;             // 首个非法字符位置（1 基），0 = 无错 [字符] / position of the first illegal character, 1 based, zero means no error [char]
END_VAR
VAR
    eState          : E_DL_StrToDintState;   // 解析状态机当前态 / current parse state
    nLen            : INT;             // 文本长度，入口锁存一次，其后全部取自该副本 [字符] / latched text length, every later bound comes from this copy [char]
    nPos            : INT;             // 字符游标（1 基）[字符] / character cursor, 1 based [char]
    nGuard          : DINT;            // WHILE 防死锁守卫计数 [次] / loop guard counter [count]
    nDigitVal       : INT;             // 当前字符的数字值，未命中为 −1 [无量纲] / numeric value of the current character, minus one when not a digit [dimensionless]
    nDigits         : INT;             // 已接受的有效数字位数 [位] / number of accepted digits [digit]
    sChar           : STRING(1);       // 当前字符，由标准 MID 取出 [字符] / current character read with the standard MID [char]
    bNeg            : BOOL;            // 负数标志，由前导符号决定 / negative flag set by the leading sign
    bAbort          : BOOL;            // 中止标志，置位后立即退出扫描 / abort flag, the scan stops as soon as it is set
    bOverflow       : BOOL;            // 溢出标志 / overflow flag
    bSpaceIgnored   : BOOL;            // 是否忽略过空格（前导或尾随）/ whether any blank was skipped, leading or trailing
    liAcc           : LINT;            // 升位累加器 [无量纲] / widened accumulator [dimensionless]
    liNext          : LINT;            // 下一拍候选累加值，先判界再落账 [无量纲] / candidate accumulator tested before it is committed [dimensionless]
    liLimit         : LINT;            // 当前符号方向下的累加上界 [无量纲] / accumulator limit for the current sign [dimensionless]
END_VAR
VAR CONSTANT
    DL_DINT_MAX         : DINT := 2147483647;        // DINT 上界，正域累加极限 [无量纲] / DINT upper bound, the positive accumulation limit [dimensionless]
    DL_DINT_MIN         : DINT := -2147483648;       // DINT 下界，负域溢出回退值 [无量纲] / DINT lower bound, the negative saturation value [dimensionless]
    DL_LINT_MAX_DINT    : LINT := 2147483647;        // 正域 LINT 判界值 [无量纲] / positive domain limit in LINT [dimensionless]
    DL_LINT_ABS_MIN     : LINT := 2147483648;        // 负域 LINT 判界值 = |DINT_MIN|，比正域大 1 [无量纲] / negative domain limit equal to the magnitude of DINT_MIN [dimensionless]
    DL_LINT_TEN         : LINT := 10;                // 十进制进位基数 [无量纲] / decimal radix [dimensionless]
    DL_STR_MAXLEN       : INT := 255;                // 文本长度上限 [字符] / text length upper bound [char]
    DL_STR_GUARD_MAX    : DINT := 600;               // 守卫上限，须大于 255 + 2 次不推进状态 / guard limit, larger than the length plus two non advancing states
    DL_STR_ONE          : INT := 1;                  // 单位哨兵 [无量纲] / unity sentinel [dimensionless]
    DL_STR_BLANK        : STRING(1) := ' ';          // 空格字符，前导与尾随都按它判 [字符] / blank character used for both ends [char]
    DL_STR_DIGITS       : STRING := '0123456789';    // 数字字符表，FIND 命中位置 − 1 即数字值 [字符] / digit table, the FIND position minus one is the value [char]
    DL_ERR_NONE         : UDINT := 16#0000_0000;     // 无故障 / no error
END_VAR

// 段 1｜返回值与错误状态预置 / segment 1, preset the return value and the error state
FC_DL_StringToDint := 0;                    // 故障缺省返回 0 / fault default returns zero
eErr           := DL_ERR_NONE;              // 预置无错误 / preset no error
bError         := FALSE;                    // 预置无故障 / preset no fault
bValid         := FALSE;                    // 预置结果不可用 / preset unusable
nErrPos        := 0;                        // 0 表示无错 / zero means no error
eState         := E_DL_StrToDintState.eLeadSpace;   // 起始态为前导空格态 / start in the leading blank state
nLen           := LEN(sIn);                 // 长度只锁存一次，禁循环内重复 LEN / latch the length once, never call LEN again in the loop
nPos           := DL_STR_ONE;               // 游标从 1 开始（MID 为 1 基）/ the cursor starts at one because MID is one based
nGuard         := 0;                        // 守卫清零 / clear the guard
nDigits        := 0;                        // 有效位数清零 / clear the digit count
nDigitVal      := 0;                        // 数字值清零 / clear the digit value
bNeg           := FALSE;                    // 预置正数 / preset positive
bAbort         := FALSE;                    // 预置不中止 / preset no abort
bOverflow      := FALSE;                    // 预置无溢出 / preset no overflow
bSpaceIgnored  := FALSE;                    // 预置未忽略空格 / preset no blank skipped
liAcc          := 0;                        // 累加器清零 / clear the accumulator
liNext         := 0;                        // 候选值清零 / clear the candidate
liLimit        := DL_LINT_MAX_DINT;         // 缺省按正域判界 / default to the positive limit
sChar          := '';                       // 字符缓冲清空 / clear the character buffer

// 段 2｜逐字符状态机：四态推进，ELSE 兜底拦非法状态 / segment 2, four state machine with an ELSE backstop
WHILE (nPos <= nLen) AND (NOT bAbort) AND (nGuard <= DL_STR_GUARD_MAX) DO
    sChar := MID(sIn, DL_STR_ONE, nPos);    // 取当前位置的一个字符 / take one character at the current position
    CASE eState OF
        E_DL_StrToDintState.eLeadSpace :
            IF sChar = DL_STR_BLANK THEN
                bSpaceIgnored := TRUE;                  // 前导空格已忽略 / a leading blank was skipped
                nPos := nPos + DL_STR_ONE;              // 前进一格 / advance one position
            ELSE
                eState := E_DL_StrToDintState.eSign;    // 转符号态，本拍不消费字符，下一轮重取同一字符 / move to the sign state without consuming this character
            END_IF

        E_DL_StrToDintState.eSign :
            IF (sChar = '+') OR (sChar = '-') THEN
                IF NOT bAllowSign THEN
                    eErr   := 16#0001_038C;             // 不允许符号却出现符号（故障级）/ a sign appeared although it is forbidden
                    bError := TRUE;                     // 置故障标志 / raise the fault flag
                    nErrPos := nPos;                    // 定位到符号位 / point at the sign
                    bAbort := TRUE;                     // 中止扫描 / abort the scan
                ELSE
                    bNeg := (sChar = '-');              // 负号判定 / detect the minus sign
                    IF bNeg THEN
                        liLimit := DL_LINT_ABS_MIN;     // 负域上界比正域大 1 / the negative limit is one larger
                    ELSE
                        liLimit := DL_LINT_MAX_DINT;    // 正域上界 / positive domain limit
                    END_IF
                    nPos   := nPos + DL_STR_ONE;        // 消费符号 / consume the sign
                    eState := E_DL_StrToDintState.eDigits;   // 转数字态 / move to the digit state
                END_IF
            ELSE
                eState := E_DL_StrToDintState.eDigits;  // 无符号直接进数字态 / no sign, go straight to the digits
            END_IF

        E_DL_StrToDintState.eDigits :
            IF sChar = DL_STR_BLANK THEN
                bSpaceIgnored := TRUE;                  // 尾随空格开始 / the trailing blanks begin
                eState := E_DL_StrToDintState.eDone;    // 转结束态，余下只允许空格 / move to done, only blanks may follow
                nPos   := nPos + DL_STR_ONE;            // 前进一格 / advance one position
            ELSE
                nDigitVal := FIND(DL_STR_DIGITS, sChar) - DL_STR_ONE;   // 命中 0~9，未命中 −1 / zero to nine when found, minus one otherwise
                IF nDigitVal < 0 THEN
                    eErr    := 16#0001_038C;            // 非法字符（故障级）/ illegal character, fault level
                    bError  := TRUE;                    // 置故障标志 / raise the fault flag
                    nErrPos := nPos;                    // 定位到首个非法字符 / point at the first illegal character
                    bAbort  := TRUE;                    // 中止扫描 / abort the scan
                ELSE
                    liNext := liAcc * DL_LINT_TEN + INT_TO_LINT(nDigitVal);   // 先算候选值 / compute the candidate first
                    IF liNext > liLimit THEN
                        bOverflow := TRUE;              // 越界即溢出，不落账 / beyond the limit means overflow, not committed
                        nErrPos   := nPos;              // 溢出位也必须定位，否则 nErrPos = 0 会被读成「无错」/ locate the overflowing digit, zero would read as no error
                        bAbort    := TRUE;              // 中止扫描 / abort the scan
                    ELSE
                        liAcc   := liNext;              // 落账 / commit
                        nDigits := nDigits + DL_STR_ONE;   // 有效位加一 / one more digit accepted
                        nPos    := nPos + DL_STR_ONE;   // 前进一格 / advance one position
                    END_IF
                    IF nPos > nLen THEN
                        eState := E_DL_StrToDintState.eDone;   // 已到串尾，转结束态 / reached the end, move to done
                    END_IF
                END_IF
            END_IF

        E_DL_StrToDintState.eDone :
            IF sChar = DL_STR_BLANK THEN
                bSpaceIgnored := TRUE;                  // 尾随空格继续忽略 / keep skipping the trailing blanks
                nPos := nPos + DL_STR_ONE;              // 前进一格 / advance one position
            ELSE
                eErr    := 16#0001_038C;                // 尾随非法字符（故障级）/ illegal trailing character, fault level
                bError  := TRUE;                        // 置故障标志 / raise the fault flag
                nErrPos := nPos;                        // 定位 / point at the position
                bAbort  := TRUE;                        // 中止扫描 / abort the scan
            END_IF

    ELSE
        // 非法状态兜底：枚举被外部改写或内存损伤，一律按「输入不可解析」处置（R90：不新占码位）
        eState   := E_DL_StrToDintState.eDone;          // 强制回已知态 / force back to a known state
        eErr     := 16#0001_038C;                      // 复用非法字符码 / reuse the illegal character code
        bError   := TRUE;                              // 置故障标志 / raise the fault flag
        nErrPos  := nPos;                              // 定位当前位 / point at the current position
        bAbort   := TRUE;                              // 中止扫描 / abort the scan
    END_CASE
    nGuard := nGuard + 1;                              // 守卫递增 / increment the guard
END_WHILE

// 段 3｜守卫复检：理论不可达（长度 ≤ 255，不推进状态最多 2 次）/ segment 3, guard re-check, unreachable in theory
IF nGuard > DL_STR_GUARD_MAX THEN
    FC_DL_StringToDint := 0;        // 不给可疑结果 / never emit a suspicious result
    eErr   := 16#0001_038C;         // 扫描失控按不可解析处置 / a runaway scan is treated as unparsable
    bError := TRUE;                 // 置故障标志 / raise the fault flag
    nErrPos := nPos;                // 定位 / point at the current position
    RETURN;                         // bValid 保持 FALSE / bValid stays FALSE
END_IF

// 段 4｜非法/溢出已中止：直接出口（故障行为已在扫描中定性）/ segment 4, exit when the scan was aborted
IF bAbort THEN
    IF bOverflow THEN
        IF bNeg THEN
            FC_DL_StringToDint := DL_DINT_MIN;   // 负域夹到下界 / saturate to the negative bound
        ELSE
            FC_DL_StringToDint := DL_DINT_MAX;   // 正域夹到上界 / saturate to the positive bound
        END_IF
        eErr := 16#0001_038B;        // 溢出已夹边界（故障级）/ overflow saturated, fault level
        bError := TRUE;              // 故障码配对置位（R101 配对，R41 P0-3 补齐）/ pair the fault flag with the fault code
    ELSE
        FC_DL_StringToDint := 0;     // 语法错误返回 0 / a syntax error returns zero
    END_IF
    RETURN;                          // bValid 保持 FALSE / bValid stays FALSE
END_IF

// 段 5｜空串或仅符号闸 / segment 5, empty string or sign-only gate
IF nDigits = 0 THEN
    FC_DL_StringToDint := 0;         // 无有效数字返回 0 / no digit at all, return zero
    eErr    := 16#0001_038A;         // 空串或仅符号（故障级）/ empty or sign only, fault level
    bError  := TRUE;                 // 置故障标志 / raise the fault flag
    nErrPos := nLen + DL_STR_ONE;    // 指向「串尾后一位」，与库内同族口径一致 / point past the end, consistent with the sibling component
    RETURN;                          // bValid 保持 FALSE / bValid stays FALSE
END_IF

// 段 6｜符号落定（下界情形在 LINT 域取负不会回绕）/ segment 6, apply the sign, negating inside LINT never wraps
IF bNeg THEN
    FC_DL_StringToDint := LINT_TO_DINT(-liAcc);   // 负域已在判界时放宽到 2147483648，故 DINT_MIN 可表达 / the limit was relaxed, so DINT_MIN is representable
ELSE
    FC_DL_StringToDint := LINT_TO_DINT(liAcc);    // 正域 / positive domain
END_IF

// 段 7｜空格提示与出口 / segment 7, blank hint and exit
IF bSpaceIgnored THEN
    eErr := 16#0001_0448;            // 前后空格已忽略（信息级，不置 bError）/ blanks ignored, info level
END_IF
bValid := TRUE;                      // 结果可用 / the result is usable
END_FUNCTION
